  movel([0.353341, -1.417894, -2.538259, -0.756236, 1.570796, 1.924137],accel_mss,speed_ms,0,blend_radius_m)
  movel([0.350688, -1.416056, -2.539657, -0.756676, 1.570796, 1.921484],accel_mss,speed_ms,0,blend_radius_m)
  movel([0.348186, -1.414065, -2.541166, -0.757158, 1.570796, 1.918982],accel_mss,speed_ms,0,blend_radius_m)
  movel([0.345836, -1.411923, -2.542783, -0.757683, 1.570796, 1.916633],accel_mss,speed_ms,0,blend_radius_m)
  movel([0.343651, -1.409630, -2.544506, -0.758253, 1.570796, 1.914447],accel_mss,speed_ms,0,blend_radius_m)
  movel([0.342913, -1.408723, -2.545186, -0.758481, 1.570796, 1.913709],accel_mss,speed_ms,0,blend_radius_m)
  movel([0.342382, -1.407674, -2.545970, -0.758745, 1.570796, 1.913178],accel_mss,speed_ms,0,blend_radius_m)
  movel([0.342236, -1.406961, -2.546502, -0.758926, 1.570796, 1.913032],accel_mss,speed_ms,0,blend_radius_m)
  movel([0.342196, -1.406201, -2.547068, -0.759119, 1.570796, 1.912992],accel_mss,speed_ms,0,blend_radius_m)
  movel([0.342303, -1.404603, -2.548257, -0.759529, 1.570796, 1.913100],accel_mss,speed_ms,0,blend_radius_m)
  movel([0.343314, -1.398696, -2.552617, -0.761077, 1.570796, 1.914110],accel_mss,speed_ms,0,blend_radius_m)
  movel([0.343428, -1.397065, -2.553812, -0.761513, 1.570796, 1.914224],accel_mss,speed_ms,0,blend_radius_m)
  movel([0.343321, -1.395654, -2.554842, -0.761893, 1.570796, 1.914117],accel_mss,speed_ms,0,blend_radius_m)
  movel([0.343156, -1.395078, -2.555262, -0.762049, 1.570796, 1.913953],accel_mss,speed_ms,0,blend_radius_m)
  movel([0.342904, -1.394608, -2.555604, -0.762177, 1.570796, 1.913701],accel_mss,speed_ms,0,blend_radius_m)
  movel([0.342554, -1.394267, -2.555852, -0.762270, 1.570796, 1.913350],accel_mss,speed_ms,0,blend_radius_m)
  movel([0.342095, -1.394069, -2.555996, -0.762324, 1.570796, 1.912892],accel_mss,speed_ms,0,blend_radius_m)
  movel([0.341153, -1.393966, -2.556071, -0.762352, 1.570796, 1.911950],accel_mss,speed_ms,0,blend_radius_m)
  movel([0.340728, -1.393866, -2.556143, -0.762379, 1.570796, 1.911524],accel_mss,speed_ms,0,blend_radius_m)
  movel([0.340432, -1.393631, -2.556314, -0.762444, 1.570796, 1.911229],accel_mss,speed_ms,0,blend_radius_m)
  movel([0.340359, -1.393040, -2.556743, -0.762606, 1.570796, 1.911155],accel_mss,speed_ms,0,blend_radius_m)
  movel([0.340573, -1.392339, -2.557251, -0.762798, 1.570796, 1.911370],accel_mss,speed_ms,0,blend_radius_m)
  movel([0.341367, -1.390085, -2.558881, -0.763423, 1.570796, 1.912163],accel_mss,speed_ms,0,blend_radius_m)
  movel([0.342003, -1.387856, -2.560485, -0.764048, 1.570796, 1.912799],accel_mss,speed_ms,0,blend_radius_m)
  movel([0.342890, -1.383456, -2.563631, -0.765302, 1.570796, 1.913686],accel_mss,speed_ms,0,blend_radius_m)
  movel([0.343413, -1.379085, -2.566728, -0.766576, 1.570796, 1.914210],accel_mss,speed_ms,0,blend_radius_m)
  movel([0.343750, -1.374694, -2.569812, -0.767883, 1.570796, 1.914546],accel_mss,speed_ms,0,blend_radius_m)
  speed_ms = 0.005
  movel([0.343750, -1.366094, -2.565773, -0.780522, 1.570796, 1.914546],accel_mss,speed_ms,0,blend_radius_m)
  speed_ms = 0.040
  movel([0.339869, -1.373054, -2.560934, -0.778400, 1.570796, 1.910666],accel_mss,speed_ms,0,blend_radius_m)
  speed_ms = 0.005
  movel([0.339869, -1.381608, -2.564943, -0.765837, 1.570796, 1.910666],accel_mss,speed_ms,0,blend_radius_m)
  speed_ms = 0.025
  movel([0.337589, -1.386297, -2.561603, -0.764489, 1.570796, 1.908385],accel_mss,speed_ms,0,blend_radius_m)
  movel([0.336311, -1.388619, -2.559937, -0.763833, 1.570796, 1.907108],accel_mss,speed_ms,0,blend_radius_m)
  movel([0.334950, -1.390919, -2.558279, -0.763191, 1.570796, 1.905746],accel_mss,speed_ms,0,blend_radius_m)
  movel([0.333977, -1.389868, -2.559037, -0.763483, 1.570796, 1.904774],accel_mss,speed_ms,0,blend_radius_m)
  movel([0.333786, -1.389712, -2.559150, -0.763527, 1.570796, 1.904582],accel_mss,speed_ms,0,blend_radius_m)
  movel([0.333516, -1.389690, -2.559166, -0.763533, 1.570796, 1.904313],accel_mss,speed_ms,0,blend_radius_m)
  movel([0.333217, -1.389876, -2.559032, -0.763481, 1.570796, 1.904013],accel_mss,speed_ms,0,blend_radius_m)
  movel([0.332976, -1.390157, -2.558829, -0.763403, 1.570796, 1.903772],accel_mss,speed_ms,0,blend_radius_m)
  movel([0.331482, -1.391896, -2.557572, -0.762921, 1.570796, 1.902279],accel_mss,speed_ms,0,blend_radius_m)
  movel([0.329770, -1.393485, -2.556421, -0.762484, 1.570796, 1.900566],accel_mss,speed_ms,0,blend_radius_m)
  movel([0.329322, -1.393797, -2.556193, -0.762398, 1.570796, 1.900118],accel_mss,speed_ms,0,blend_radius_m)
  movel([0.328892, -1.393891, -2.556126, -0.762373, 1.570796, 1.899688],accel_mss,speed_ms,0,blend_radius_m)
  movel([0.328696, -1.393685, -2.556275, -0.762429, 1.570796, 1.899492],accel_mss,speed_ms,0,blend_radius_m)
  movel([0.328675, -1.393350, -2.556518, -0.762521, 1.570796, 1.899472],accel_mss,speed_ms,0,blend_radius_m)
  movel([0.328990, -1.391182, -2.558089, -0.763118, 1.570796, 1.899786],accel_mss,speed_ms,0,blend_radius_m)
  movel([0.329681, -1.388937, -2.559708, -0.763744, 1.570796, 1.900478],accel_mss,speed_ms,0,blend_radius_m)
  speed_ms = 0.005
  movel([0.329681, -1.380434, -2.555730, -0.776225, 1.570796, 1.900478],accel_mss,speed_ms,0,blend_radius_m)
  speed_ms = 0.040
  movel([0.332271, -1.385014, -2.552462, -0.774913, 1.570796, 1.903067],accel_mss,speed_ms,0,blend_radius_m)
  speed_ms = 0.005
  movel([0.332271, -1.393486, -2.556420, -0.762483, 1.570796, 1.903067],accel_mss,speed_ms,0,blend_radius_m)
  speed_ms = 0.025
  movel([0.331292, -1.396772, -2.554026, -0.761592, 1.570796, 1.902088],accel_mss,speed_ms,0,blend_radius_m)
  movel([0.330631, -1.398425, -2.552816, -0.761149, 1.570796, 1.901428],accel_mss,speed_ms,0,blend_radius_m)
  movel([0.328994, -1.401710, -2.550398, -0.760281, 1.570796, 1.899790],accel_mss,speed_ms,0,blend_radius_m)
  movel([0.328023, -1.403329, -2.549201, -0.759859, 1.570796, 1.898819],accel_mss,speed_ms,0,blend_radius_m)
  movel([0.325798, -1.406488, -2.546855, -0.759046, 1.570796, 1.896594],accel_mss,speed_ms,0,blend_radius_m)
  movel([0.326216, -1.405393, -2.547669, -0.759326, 1.570796, 1.897012],accel_mss,speed_ms,0,blend_radius_m)
  movel([0.326316, -1.404349, -2.548445, -0.759595, 1.570796, 1.897112],accel_mss,speed_ms,0,blend_radius_m)
  movel([0.326100, -1.403427, -2.549128, -0.759833, 1.570796, 1.896896],accel_mss,speed_ms,0,blend_radius_m)
  movel([0.325568, -1.402702, -2.549666, -0.760022, 1.570796, 1.896365],accel_mss,speed_ms,0,blend_radius_m)
  speed_ms = 0.005
  movel([0.325568, -1.394294, -2.545747, -0.772348, 1.570796, 1.896365],accel_mss,speed_ms,0,blend_radius_m)
  speed_ms = 0.040
  movel([0.312695, -1.397176, -2.543637, -0.771576, 1.570796, 1.883492],accel_mss,speed_ms,0,blend_radius_m)
  speed_ms = 0.005
  movel([0.312695, -1.405564, -2.547543, -0.759283, 1.570796, 1.883492],accel_mss,speed_ms,0,blend_radius_m)
  speed_ms = 0.025
  movel([0.310320, -1.407416, -2.546163, -0.758811, 1.570796, 1.881117],accel_mss,speed_ms,0,blend_radius_m)
  movel([0.307808, -1.409042, -2.544946, -0.758400, 1.570796, 1.878604],accel_mss,speed_ms,0,blend_radius_m)
  movel([0.305202, -1.410422, -2.543912, -0.758055, 1.570796, 1.875999],accel_mss,speed_ms,0,blend_radius_m)
  movel([0.302547, -1.411527, -2.543081, -0.757781, 1.570796, 1.873344],accel_mss,speed_ms,0,blend_radius_m)
  movel([0.303286, -1.410545, -2.543819, -0.758025, 1.570796, 1.874082],accel_mss,speed_ms,0,blend_radius_m)
  movel([0.303859, -1.409585, -2.544540, -0.758264, 1.570796, 1.874656],accel_mss,speed_ms,0,blend_radius_m)
  movel([0.304225, -1.408734, -2.545177, -0.758478, 1.570796, 1.875021],accel_mss,speed_ms,0,blend_radius_m)
  movel([0.304341, -1.408081, -2.545666, -0.758642, 1.570796, 1.875137],accel_mss,speed_ms,0,blend_radius_m)
  movel([0.304161, -1.407717, -2.545938, -0.758734, 1.570796, 1.874957],accel_mss,speed_ms,0,blend_radius_m)
  movel([0.303948, -1.407671, -2.545972, -0.758746, 1.570796, 1.874744],accel_mss,speed_ms,0,blend_radius_m)
  movel([0.303642, -1.407729, -2.545928, -0.758731, 1.570796, 1.874438],accel_mss,speed_ms,0,blend_radius_m)
  movel([0.302742, -1.408211, -2.545569, -0.758610, 1.570796, 1.873539],accel_mss,speed_ms,0,blend_radius_m)
  movel([0.300391, -1.410083, -2.544167, -0.758140, 1.570796, 1.871188],accel_mss,speed_ms,0,blend_radius_m)
  movel([0.299301, -1.410867, -2.543577, -0.757945, 1.570796, 1.870098],accel_mss,speed_ms,0,blend_radius_m)
  movel([0.296993, -1.412235, -2.542548, -0.757606, 1.570796, 1.867789],accel_mss,speed_ms,0,blend_radius_m)
  movel([0.295802, -1.412800, -2.542122, -0.757467, 1.570796, 1.866599],accel_mss,speed_ms,0,blend_radius_m)
  movel([0.294607, -1.413268, -2.541769, -0.757352, 1.570796, 1.865403],accel_mss,speed_ms,0,blend_radius_m)
  movel([0.293418, -1.413635, -2.541492, -0.757263, 1.570796, 1.864215],accel_mss,speed_ms,0,blend_radius_m)
  movel([0.292256, -1.413884, -2.541303, -0.757202, 1.570796, 1.863052],accel_mss,speed_ms,0,blend_radius_m)
  movel([0.293826, -1.412474, -2.542367, -0.757547, 1.570796, 1.864623],accel_mss,speed_ms,0,blend_radius_m)
  movel([0.295363, -1.411029, -2.543456, -0.757904, 1.570796, 1.866160],accel_mss,speed_ms,0,blend_radius_m)
  movel([0.296110, -1.409980, -2.544243, -0.758165, 1.570796, 1.866906],accel_mss,speed_ms,0,blend_radius_m)
  movel([0.296586, -1.408893, -2.545058, -0.758438, 1.570796, 1.867383],accel_mss,speed_ms,0,blend_radius_m)
  movel([0.296599, -1.408490, -2.545359, -0.758539, 1.570796, 1.867396],accel_mss,speed_ms,0,blend_radius_m)
  movel([0.296393, -1.408265, -2.545528, -0.758596, 1.570796, 1.867190],accel_mss,speed_ms,0,blend_radius_m)
  movel([0.295922, -1.408281, -2.545516, -0.758592, 1.570796, 1.866719],accel_mss,speed_ms,0,blend_radius_m)
  movel([0.295135, -1.408602, -2.545276, -0.758511, 1.570796, 1.865931],accel_mss,speed_ms,0,blend_radius_m)
  movel([0.290915, -1.410859, -2.543584, -0.757947, 1.570796, 1.861712],accel_mss,speed_ms,0,blend_radius_m)
  movel([0.288820, -1.411752, -2.542911, -0.757725, 1.570796, 1.859616],accel_mss,speed_ms,0,blend_radius_m)
  movel([0.287788, -1.412048, -2.542689, -0.757652, 1.570796, 1.858584],accel_mss,speed_ms,0,blend_radius_m)
  movel([0.286768, -1.412208, -2.542568, -0.757613, 1.570796, 1.857565],accel_mss,speed_ms,0,blend_radius_m)
  speed_ms = 0.005
  movel([0.286768, -1.403867, -2.538690, -0.769831, 1.570796, 1.857565],accel_mss,speed_ms,0,blend_radius_m)
  speed_ms = 0.040
  movel([0.307123, -1.384967, -2.552495, -0.774927, 1.570796, 1.877919],accel_mss,speed_ms,0,blend_radius_m)
  speed_ms = 0.005
  movel([0.307123, -1.393440, -2.556453, -0.762496, 1.570796, 1.877919],accel_mss,speed_ms,0,blend_radius_m)
  speed_ms = 0.025
  movel([0.307349, -1.392012, -2.557488, -0.762888, 1.570796, 1.878145],accel_mss,speed_ms,0,blend_radius_m)
  movel([0.307875, -1.390552, -2.558544, -0.763293, 1.570796, 1.878671],accel_mss,speed_ms,0,blend_radius_m)
  movel([0.308665, -1.389081, -2.559605, -0.763704, 1.570796, 1.879461],accel_mss,speed_ms,0,blend_radius_m)
  movel([0.309681, -1.387631, -2.560646, -0.764111, 1.570796, 1.880477],accel_mss,speed_ms,0,blend_radius_m)
  movel([0.310891, -1.386226, -2.561654, -0.764509, 1.570796, 1.881688],accel_mss,speed_ms,0,blend_radius_m)
  movel([0.312255, -1.384897, -2.562603, -0.764888, 1.570796, 1.883051],accel_mss,speed_ms,0,blend_radius_m)
  movel([0.313741, -1.383669, -2.563479, -0.765241, 1.570796, 1.884537],accel_mss,speed_ms,0,blend_radius_m)
  movel([0.315307, -1.382571, -2.564260, -0.765558, 1.570796, 1.886103],accel_mss,speed_ms,0,blend_radius_m)
  movel([0.317303, -1.381387, -2.565100, -0.765902, 1.570796, 1.888099],accel_mss,speed_ms,0,blend_radius_m)
  movel([0.321349, -1.379143, -2.566687, -0.766559, 1.570796, 1.892145],accel_mss,speed_ms,0,blend_radius_m)
  movel([0.323312, -1.377877, -2.567579, -0.766933, 1.570796, 1.894108],accel_mss,speed_ms,0,blend_radius_m)
  movel([0.325159, -1.376347, -2.568654, -0.767388, 1.570796, 1.895955],accel_mss,speed_ms,0,blend_radius_m)
  movel([0.325987, -1.375488, -2.569256, -0.767645, 1.570796, 1.896784],accel_mss,speed_ms,0,blend_radius_m)
  movel([0.326715, -1.374590, -2.569885, -0.767914, 1.570796, 1.897511],accel_mss,speed_ms,0,blend_radius_m)
  movel([0.327314, -1.373670, -2.570527, -0.768192, 1.570796, 1.898111],accel_mss,speed_ms,0,blend_radius_m)
  movel([0.327760, -1.372746, -2.571172, -0.768472, 1.570796, 1.898557],accel_mss,speed_ms,0,blend_radius_m)
  movel([0.328019, -1.371841, -2.571802, -0.768747, 1.570796, 1.898816],accel_mss,speed_ms,0,blend_radius_m)
  movel([0.328063, -1.370972, -2.572405, -0.769012, 1.570796, 1.898860],accel_mss,speed_ms,0,blend_radius_m)
  speed_ms = 0.005
  movel([0.328063, -1.362347, -2.568349, -0.781693, 1.570796, 1.898860],accel_mss,speed_ms,0,blend_radius_m)
  speed_ms = 0.040
  movel([0.327969, -1.355374, -2.573093, -0.783923, 1.570796, 1.898765],accel_mss,speed_ms,0,blend_radius_m)
  speed_ms = 0.005
  movel([0.327969, -1.364044, -2.577178, -0.771166, 1.570796, 1.898765],accel_mss,speed_ms,0,blend_radius_m)
  speed_ms = 0.025
  movel([0.325748, -1.369382, -2.573506, -0.769501, 1.570796, 1.896545],accel_mss,speed_ms,0,blend_radius_m)
  movel([0.325014, -1.370536, -2.572707, -0.769146, 1.570796, 1.895810],accel_mss,speed_ms,0,blend_radius_m)
  movel([0.323980, -1.371546, -2.572006, -0.768837, 1.570796, 1.894777],accel_mss,speed_ms,0,blend_radius_m)
  movel([0.322764, -1.372368, -2.571435, -0.768586, 1.570796, 1.893560],accel_mss,speed_ms,0,blend_radius_m)
  movel([0.318705, -1.374593, -2.569882, -0.767913, 1.570796, 1.889501],accel_mss,speed_ms,0,blend_radius_m)
  movel([0.317313, -1.375524, -2.569231, -0.767634, 1.570796, 1.888110],accel_mss,speed_ms,0,blend_radius_m)
  movel([0.315981, -1.376546, -2.568514, -0.767328, 1.570796, 1.886777],accel_mss,speed_ms,0,blend_radius_m)
  movel([0.314719, -1.377645, -2.567743, -0.767002, 1.570796, 1.885516],accel_mss,speed_ms,0,blend_radius_m)
  movel([0.313629, -1.378816, -2.566918, -0.766655, 1.570796, 1.884425],accel_mss,speed_ms,0,blend_radius_m)
  movel([0.312677, -1.380053, -2.566044, -0.766292, 1.570796, 1.883473],accel_mss,speed_ms,0,blend_radius_m)
  movel([0.311739, -1.381287, -2.565171, -0.765931, 1.570796, 1.882535],accel_mss,speed_ms,0,blend_radius_m)
  movel([0.310692, -1.382453, -2.564344, -0.765592, 1.570796, 1.881488],accel_mss,speed_ms,0,blend_radius_m)
  movel([0.310217, -1.379416, -2.566495, -0.766479, 1.570796, 1.881013],accel_mss,speed_ms,0,blend_radius_m)
  movel([0.310427, -1.378523, -2.567124, -0.766742, 1.570796, 1.881223],accel_mss,speed_ms,0,blend_radius_m)
  movel([0.310784, -1.377639, -2.567747, -0.767003, 1.570796, 1.881580],accel_mss,speed_ms,0,blend_radius_m)
  movel([0.311287, -1.376761, -2.568364, -0.767264, 1.570796, 1.882083],accel_mss,speed_ms,0,blend_radius_m)
  movel([0.311945, -1.375885, -2.568978, -0.767526, 1.570796, 1.882741],accel_mss,speed_ms,0,blend_radius_m)
  movel([0.313120, -1.374783, -2.569750, -0.767856, 1.570796, 1.883917],accel_mss,speed_ms,0,blend_radius_m)
  movel([0.314797, -1.373557, -2.570606, -0.768226, 1.570796, 1.885594],accel_mss,speed_ms,0,blend_radius_m)
  movel([0.318871, -1.370934, -2.572431, -0.769024, 1.570796, 1.889668],accel_mss,speed_ms,0,blend_radius_m)
  movel([0.320876, -1.369641, -2.573327, -0.769421, 1.570796, 1.891672],accel_mss,speed_ms,0,blend_radius_m)
  movel([0.322594, -1.368424, -2.574168, -0.769796, 1.570796, 1.893391],accel_mss,speed_ms,0,blend_radius_m)
  movel([0.323827, -1.367340, -2.574916, -0.770133, 1.570796, 1.894624],accel_mss,speed_ms,0,blend_radius_m)
  movel([0.324201, -1.366860, -2.575247, -0.770283, 1.570796, 1.894997],accel_mss,speed_ms,0,blend_radius_m)
  movel([0.324377, -1.366430, -2.575542, -0.770417, 1.570796, 1.895173],accel_mss,speed_ms,0,blend_radius_m)
  speed_ms = 0.005
  movel([0.324377, -1.357775, -2.571467, -0.783147, 1.570796, 1.895173],accel_mss,speed_ms,0,blend_radius_m)
  speed_ms = 0.040
  movel([0.317644, -1.355816, -2.572794, -0.783779, 1.570796, 1.888440],accel_mss,speed_ms,0,blend_radius_m)
  speed_ms = 0.005
  movel([0.317644, -1.364484, -2.576878, -0.771028, 1.570796, 1.888440],accel_mss,speed_ms,0,blend_radius_m)
  speed_ms = 0.025
  movel([0.316995, -1.364280, -2.577017, -0.771092, 1.570796, 1.887792],accel_mss,speed_ms,0,blend_radius_m)
  movel([0.316480, -1.363934, -2.577254, -0.771201, 1.570796, 1.887276],accel_mss,speed_ms,0,blend_radius_m)
  movel([0.315783, -1.362916, -2.577950, -0.771524, 1.570796, 1.886579],accel_mss,speed_ms,0,blend_radius_m)
  movel([0.315427, -1.361607, -2.578842, -0.771940, 1.570796, 1.886224],accel_mss,speed_ms,0,blend_radius_m)
  movel([0.315292, -1.360185, -2.579809, -0.772396, 1.570796, 1.886089],accel_mss,speed_ms,0,blend_radius_m)
  movel([0.315340, -1.359638, -2.580180, -0.772572, 1.570796, 1.886136],accel_mss,speed_ms,0,blend_radius_m)
  movel([0.315896, -1.358775, -2.580764, -0.772850, 1.570796, 1.886692],accel_mss,speed_ms,0,blend_radius_m)
  movel([0.317769, -1.356422, -2.582353, -0.773614, 1.570796, 1.888565],accel_mss,speed_ms,0,blend_radius_m)
  movel([0.321286, -1.351596, -2.585588, -0.775206, 1.570796, 1.892083],accel_mss,speed_ms,0,blend_radius_m)
  movel([0.322923, -1.349133, -2.587226, -0.776031, 1.570796, 1.893720],accel_mss,speed_ms,0,blend_radius_m)
  speed_ms = 0.005
  movel([0.322923, -1.340366, -2.583075, -0.788949, 1.570796, 1.893720],accel_mss,speed_ms,0,blend_radius_m)
  speed_ms = 0.040
  movel([0.318249, -1.341582, -2.582277, -0.788530, 1.570796, 1.889045],accel_mss,speed_ms,0,blend_radius_m)
  speed_ms = 0.005
  movel([0.318249, -1.350341, -2.586423, -0.775625, 1.570796, 1.889045],accel_mss,speed_ms,0,blend_radius_m)
  speed_ms = 0.025
  movel([0.317404, -1.351859, -2.585412, -0.775118, 1.570796, 1.888200],accel_mss,speed_ms,0,blend_radius_m)
  movel([0.316388, -1.353339, -2.584423, -0.774627, 1.570796, 1.887185],accel_mss,speed_ms,0,blend_radius_m)
  movel([0.315173, -1.354678, -2.583525, -0.774186, 1.570796, 1.885969],accel_mss,speed_ms,0,blend_radius_m)
  movel([0.314479, -1.355266, -2.583131, -0.773992, 1.570796, 1.885275],accel_mss,speed_ms,0,blend_radius_m)
  movel([0.312991, -1.356296, -2.582438, -0.773655, 1.570796, 1.883787],accel_mss,speed_ms,0,blend_radius_m)
  movel([0.312589, -1.356891, -2.582037, -0.773461, 1.570796, 1.883385],accel_mss,speed_ms,0,blend_radius_m)
  movel([0.310058, -1.361595, -2.578850, -0.771944, 1.570796, 1.880854],accel_mss,speed_ms,0,blend_radius_m)
  movel([0.309827, -1.362051, -2.578539, -0.771798, 1.570796, 1.880623],accel_mss,speed_ms,0,blend_radius_m)
  movel([0.309727, -1.362487, -2.578242, -0.771660, 1.570796, 1.880524],accel_mss,speed_ms,0,blend_radius_m)
  movel([0.309968, -1.362959, -2.577920, -0.771510, 1.570796, 1.880764],accel_mss,speed_ms,0,blend_radius_m)
  movel([0.310464, -1.363243, -2.577726, -0.771420, 1.570796, 1.881260],accel_mss,speed_ms,0,blend_radius_m)
  movel([0.311933, -1.363994, -2.577213, -0.771182, 1.570796, 1.882730],accel_mss,speed_ms,0,blend_radius_m)
  movel([0.313243, -1.364912, -2.576584, -0.770893, 1.570796, 1.884039],accel_mss,speed_ms,0,blend_radius_m)
  movel([0.314279, -1.366052, -2.575802, -0.770535, 1.570796, 1.885076],accel_mss,speed_ms,0,blend_radius_m)
  movel([0.314920, -1.367474, -2.574824, -0.770091, 1.570796, 1.885717],accel_mss,speed_ms,0,blend_radius_m)
  speed_ms = 0.005
  movel([0.314920, -1.358825, -2.570753, -0.782811, 1.570796, 1.885717],accel_mss,speed_ms,0,blend_radius_m)
  speed_ms = 0.040
  movel([0.308499, -1.370918, -2.562427, -0.779044, 1.570796, 1.879295],accel_mss,speed_ms,0,blend_radius_m)
  speed_ms = 0.005
  movel([0.308499, -1.379486, -2.566445, -0.766458, 1.570796, 1.879295],accel_mss,speed_ms,0,blend_radius_m)
  speed_ms = 0.025
  movel([0.308142, -1.379675, -2.566311, -0.766402, 1.570796, 1.878938],accel_mss,speed_ms,0,blend_radius_m)
  movel([0.307804, -1.379962, -2.566109, -0.766318, 1.570796, 1.878600],accel_mss,speed_ms,0,blend_radius_m)
  movel([0.306398, -1.381586, -2.564959, -0.765844, 1.570796, 1.877194],accel_mss,speed_ms,0,blend_radius_m)
  movel([0.306182, -1.381703, -2.564876, -0.765810, 1.570796, 1.876978],accel_mss,speed_ms,0,blend_radius_m)
  movel([0.305890, -1.381676, -2.564896, -0.765818, 1.570796, 1.876686],accel_mss,speed_ms,0,blend_radius_m)
  movel([0.305691, -1.381462, -2.565047, -0.765880, 1.570796, 1.876488],accel_mss,speed_ms,0,blend_radius_m)
  movel([0.305524, -1.380686, -2.565597, -0.766106, 1.570796, 1.876321],accel_mss,speed_ms,0,blend_radius_m)
  movel([0.305660, -1.379126, -2.566699, -0.766564, 1.570796, 1.876456],accel_mss,speed_ms,0,blend_radius_m)
  movel([0.306239, -1.377612, -2.567766, -0.767011, 1.570796, 1.877035],accel_mss,speed_ms,0,blend_radius_m)
  movel([0.307051, -1.376086, -2.568837, -0.767465, 1.570796, 1.877848],accel_mss,speed_ms,0,blend_radius_m)
  movel([0.307976, -1.374599, -2.569878, -0.767911, 1.570796, 1.878772],accel_mss,speed_ms,0,blend_radius_m)
  movel([0.309020, -1.373202, -2.570853, -0.768333, 1.570796, 1.879816],accel_mss,speed_ms,0,blend_radius_m)
  movel([0.310178, -1.371895, -2.571763, -0.768730, 1.570796, 1.880974],accel_mss,speed_ms,0,blend_radius_m)
  movel([0.311443, -1.370676, -2.572610, -0.769103, 1.570796, 1.882240],accel_mss,speed_ms,0,blend_radius_m)
  movel([0.312813, -1.369539, -2.573398, -0.769452, 1.570796, 1.883610],accel_mss,speed_ms,0,blend_radius_m)
  movel([0.314279, -1.368486, -2.574126, -0.769777, 1.570796, 1.885075],accel_mss,speed_ms,0,blend_radius_m)
  movel([0.315839, -1.367510, -2.574799, -0.770080, 1.570796, 1.886635],accel_mss,speed_ms,0,blend_radius_m)
  movel([0.317485, -1.366610, -2.575418, -0.770361, 1.570796, 1.888282],accel_mss,speed_ms,0,blend_radius_m)
  movel([0.319775, -1.365190, -2.576393, -0.770805, 1.570796, 1.890571],accel_mss,speed_ms,0,blend_radius_m)
  movel([0.322192, -1.363404, -2.577616, -0.771369, 1.570796, 1.892989],accel_mss,speed_ms,0,blend_radius_m)
  movel([0.324813, -1.361260, -2.579078, -0.772051, 1.570796, 1.895609],accel_mss,speed_ms,0,blend_radius_m)
  speed_ms = 0.005
  movel([0.324813, -1.352571, -2.574980, -0.784838, 1.570796, 1.895609],accel_mss,speed_ms,0,blend_radius_m)
  speed_ms = 0.040
  movel([0.322789, -1.352336, -2.575138, -0.784915, 1.570796, 1.893585],accel_mss,speed_ms,0,blend_radius_m)
  speed_ms = 0.005
  movel([0.322789, -1.361026, -2.579237, -0.772126, 1.570796, 1.893585],accel_mss,speed_ms,0,blend_radius_m)
  speed_ms = 0.025
  movel([0.325060, -1.357489, -2.581633, -0.773266, 1.570796, 1.895856],accel_mss,speed_ms,0,blend_radius_m)
  movel([0.327540, -1.353985, -2.583990, -0.774414, 1.570796, 1.898337],accel_mss,speed_ms,0,blend_radius_m)
  movel([0.328901, -1.352289, -2.585125, -0.774975, 1.570796, 1.899697],accel_mss,speed_ms,0,blend_radius_m)
  movel([0.330358, -1.350651, -2.586217, -0.775521, 1.570796, 1.901154],accel_mss,speed_ms,0,blend_radius_m)
  movel([0.331934, -1.349089, -2.587255, -0.776045, 1.570796, 1.902731],accel_mss,speed_ms,0,blend_radius_m)
  movel([0.333636, -1.347623, -2.588226, -0.776540, 1.570796, 1.904433],accel_mss,speed_ms,0,blend_radius_m)
  movel([0.338281, -1.344182, -2.590494, -0.777714, 1.570796, 1.909077],accel_mss,speed_ms,0,blend_radius_m)
  movel([0.340290, -1.342554, -2.591561, -0.778274, 1.570796, 1.911086],accel_mss,speed_ms,0,blend_radius_m)
  movel([0.341243, -1.341682, -2.592131, -0.778576, 1.570796, 1.912039],accel_mss,speed_ms,0,blend_radius_m)
  movel([0.342119, -1.340743, -2.592744, -0.778902, 1.570796, 1.912915],accel_mss,speed_ms,0,blend_radius_m)
  movel([0.344165, -1.337635, -2.594763, -0.779991, 1.570796, 1.914961],accel_mss,speed_ms,0,blend_radius_m)
  speed_ms = 0.005
  movel([0.344165, -1.328796, -2.590561, -0.793032, 1.570796, 1.914961],accel_mss,speed_ms,0,blend_radius_m)
  speed_ms = 0.040
  movel([0.349051, -1.321604, -2.595125, -0.795660, 1.570796, 1.919847],accel_mss,speed_ms,0,blend_radius_m)
  speed_ms = 0.005
  movel([0.349051, -1.330486, -2.599359, -0.782543, 1.570796, 1.919847],accel_mss,speed_ms,0,blend_radius_m)
  speed_ms = 0.025
  movel([0.350619, -1.327900, -2.601005, -0.783484, 1.570796, 1.921415],accel_mss,speed_ms,0,blend_radius_m)
  movel([0.351604, -1.326705, -2.601762, -0.783922, 1.570796, 1.922400],accel_mss,speed_ms,0,blend_radius_m)
  movel([0.352794, -1.325669, -2.602418, -0.784303, 1.570796, 1.923590],accel_mss,speed_ms,0,blend_radius_m)
  movel([0.353735, -1.325094, -2.602780, -0.784515, 1.570796, 1.924531],accel_mss,speed_ms,0,blend_radius_m)
  movel([0.354708, -1.324645, -2.603064, -0.784681, 1.570796, 1.925504],accel_mss,speed_ms,0,blend_radius_m)
  movel([0.356688, -1.323931, -2.603513, -0.784945, 1.570796, 1.927484],accel_mss,speed_ms,0,blend_radius_m)
  movel([0.358468, -1.323146, -2.604007, -0.785236, 1.570796, 1.929265],accel_mss,speed_ms,0,blend_radius_m)
  movel([0.359922, -1.322182, -2.604612, -0.785595, 1.570796, 1.930719],accel_mss,speed_ms,0,blend_radius_m)
  movel([0.362751, -1.319636, -2.606203, -0.786549, 1.570796, 1.933547],accel_mss,speed_ms,0,blend_radius_m)
  movel([0.363357, -1.319157, -2.606502, -0.786730, 1.570796, 1.934153],accel_mss,speed_ms,0,blend_radius_m)
  movel([0.364004, -1.318782, -2.606736, -0.786871, 1.570796, 1.934800],accel_mss,speed_ms,0,blend_radius_m)
  movel([0.365382, -1.318258, -2.607061, -0.787069, 1.570796, 1.936179],accel_mss,speed_ms,0,blend_radius_m)
  movel([0.368164, -1.317488, -2.607540, -0.787361, 1.570796, 1.938960],accel_mss,speed_ms,0,blend_radius_m)
  movel([0.371123, -1.316378, -2.608228, -0.787783, 1.570796, 1.941919],accel_mss,speed_ms,0,blend_radius_m)
  movel([0.372596, -1.315685, -2.608657, -0.788047, 1.570796, 1.943392],accel_mss,speed_ms,0,blend_radius_m)
  movel([0.374034, -1.314815, -2.609194, -0.788379, 1.570796, 1.944830],accel_mss,speed_ms,0,blend_radius_m)
  movel([0.375107, -1.313914, -2.609750, -0.788725, 1.570796, 1.945903],accel_mss,speed_ms,0,blend_radius_m)
  movel([0.375975, -1.312857, -2.610400, -0.789131, 1.570796, 1.946771],accel_mss,speed_ms,0,blend_radius_m)
  movel([0.376436, -1.311818, -2.611038, -0.789533, 1.570796, 1.947232],accel_mss,speed_ms,0,blend_radius_m)
  movel([0.376451, -1.311361, -2.611318, -0.789709, 1.570796, 1.947248],accel_mss,speed_ms,0,blend_radius_m)
  movel([0.376289, -1.310975, -2.611555, -0.789859, 1.570796, 1.947085],accel_mss,speed_ms,0,blend_radius_m)
  movel([0.375621, -1.310415, -2.611897, -0.790077, 1.570796, 1.946417],accel_mss,speed_ms,0,blend_radius_m)
  movel([0.374663, -1.310045, -2.612124, -0.790220, 1.570796, 1.945460],accel_mss,speed_ms,0,blend_radius_m)
  movel([0.373483, -1.309859, -2.612237, -0.790293, 1.570796, 1.944279],accel_mss,speed_ms,0,blend_radius_m)
  movel([0.372161, -1.309843, -2.612247, -0.790299, 1.570796, 1.942958],accel_mss,speed_ms,0,blend_radius_m)
  movel([0.370770, -1.309993, -2.612155, -0.790241, 1.570796, 1.941566],accel_mss,speed_ms,0,blend_radius_m)
  movel([0.369387, -1.310295, -2.611971, -0.790123, 1.570796, 1.940183],accel_mss,speed_ms,0,blend_radius_m)
  movel([0.368086, -1.310742, -2.611697, -0.789950, 1.570796, 1.938882],accel_mss,speed_ms,0,blend_radius_m)
  movel([0.366941, -1.311323, -2.611342, -0.789724, 1.570796, 1.937738],accel_mss,speed_ms,0,blend_radius_m)
  movel([0.365361, -1.312504, -2.610617, -0.789268, 1.570796, 1.936157],accel_mss,speed_ms,0,blend_radius_m)
  movel([0.360899, -1.316398, -2.608216, -0.787775, 1.570796, 1.931696],accel_mss,speed_ms,0,blend_radius_m)
  movel([0.357794, -1.318784, -2.606735, -0.786871, 1.570796, 1.928590],accel_mss,speed_ms,0,blend_radius_m)
  movel([0.354959, -1.320535, -2.605642, -0.786211, 1.570796, 1.925755],accel_mss,speed_ms,0,blend_radius_m)
  movel([0.353550, -1.321372, -2.605119, -0.785898, 1.570796, 1.924347],accel_mss,speed_ms,0,blend_radius_m)
  movel([0.352205, -1.322311, -2.604531, -0.785547, 1.570796, 1.923002],accel_mss,speed_ms,0,blend_radius_m)
  movel([0.350915, -1.323430, -2.603828, -0.785131, 1.570796, 1.921711],accel_mss,speed_ms,0,blend_radius_m)
  movel([0.349740, -1.324629, -2.603073, -0.784686, 1.570796, 1.920536],accel_mss,speed_ms,0,blend_radius_m)
  movel([0.348669, -1.325894, -2.602275, -0.784220, 1.570796, 1.919466],accel_mss,speed_ms,0,blend_radius_m)
  movel([0.347691, -1.327204, -2.601446, -0.783739, 1.570796, 1.918487],accel_mss,speed_ms,0,blend_radius_m)
  movel([0.345956, -1.329897, -2.599735, -0.782757, 1.570796, 1.916752],accel_mss,speed_ms,0,blend_radius_m)
  movel([0.344424, -1.332576, -2.598023, -0.781790, 1.570796, 1.915221],accel_mss,speed_ms,0,blend_radius_m)
  speed_ms = 0.005
  movel([0.344424, -1.323706, -2.593798, -0.794885, 1.570796, 1.915221],accel_mss,speed_ms,0,blend_radius_m)
  speed_ms = 0.040
  movel([0.340785, -1.325157, -2.592879, -0.794353, 1.570796, 1.911581],accel_mss,speed_ms,0,blend_radius_m)
  speed_ms = 0.005
  movel([0.340785, -1.334019, -2.597097, -0.781273, 1.570796, 1.911581],accel_mss,speed_ms,0,blend_radius_m)
  speed_ms = 0.025
  movel([0.343327, -1.329820, -2.599784, -0.782785, 1.570796, 1.914124],accel_mss,speed_ms,0,blend_radius_m)
  movel([0.344465, -1.328079, -2.600891, -0.783419, 1.570796, 1.915261],accel_mss,speed_ms,0,blend_radius_m)
  movel([0.345507, -1.326318, -2.602007, -0.784064, 1.570796, 1.916304],accel_mss,speed_ms,0,blend_radius_m)
  movel([0.346218, -1.324778, -2.602980, -0.784631, 1.570796, 1.917014],accel_mss,speed_ms,0,blend_radius_m)
  movel([0.346717, -1.323245, -2.603944, -0.785199, 1.570796, 1.917514],accel_mss,speed_ms,0,blend_radius_m)
  movel([0.346996, -1.321750, -2.604882, -0.785757, 1.570796, 1.917792],accel_mss,speed_ms,0,blend_radius_m)
  movel([0.347046, -1.320325, -2.605774, -0.786290, 1.570796, 1.917842],accel_mss,speed_ms,0,blend_radius_m)
  movel([0.347778, -1.320120, -2.605901, -0.786367, 1.570796, 1.918574],accel_mss,speed_ms,0,blend_radius_m)
  movel([0.348472, -1.320081, -2.605926, -0.786382, 1.570796, 1.919268],accel_mss,speed_ms,0,blend_radius_m)
  movel([0.349799, -1.320203, -2.605850, -0.786336, 1.570796, 1.920596],accel_mss,speed_ms,0,blend_radius_m)
  movel([0.351211, -1.320202, -2.605850, -0.786337, 1.570796, 1.922008],accel_mss,speed_ms,0,blend_radius_m)
  movel([0.351944, -1.320017, -2.605966, -0.786406, 1.570796, 1.922741],accel_mss,speed_ms,0,blend_radius_m)
  movel([0.352658, -1.319621, -2.606213, -0.786555, 1.570796, 1.923455],accel_mss,speed_ms,0,blend_radius_m)
  movel([0.360769, -1.313713, -2.609874, -0.788802, 1.570796, 1.931565],accel_mss,speed_ms,0,blend_radius_m)
  movel([0.360914, -1.312683, -2.610507, -0.789199, 1.570796, 1.931710],accel_mss,speed_ms,0,blend_radius_m)
  movel([0.360736, -1.311745, -2.611083, -0.789561, 1.570796, 1.931532],accel_mss,speed_ms,0,blend_radius_m)
  movel([0.360245, -1.310950, -2.611570, -0.789869, 1.570796, 1.931041],accel_mss,speed_ms,0,blend_radius_m)
  movel([0.359461, -1.310345, -2.611940, -0.790104, 1.570796, 1.930257],accel_mss,speed_ms,0,blend_radius_m)
  movel([0.361095, -1.310189, -2.612035, -0.790164, 1.570796, 1.931891],accel_mss,speed_ms,0,blend_radius_m)
  movel([0.362585, -1.310328, -2.611951, -0.790110, 1.570796, 1.933381],accel_mss,speed_ms,0,blend_radius_m)
  movel([0.363857, -1.310746, -2.611695, -0.789948, 1.570796, 1.934653],accel_mss,speed_ms,0,blend_radius_m)
  movel([0.364841, -1.311428, -2.611277, -0.789684, 1.570796, 1.935638],accel_mss,speed_ms,0,blend_radius_m)
  speed_ms = 0.005
  movel([0.364841, -1.302433, -2.606958, -0.802997, 1.570796, 1.935638],accel_mss,speed_ms,0,blend_radius_m)
  speed_ms = 0.040
  movel([0.366450, -1.298436, -2.609366, -0.804587, 1.570796, 1.937246],accel_mss,speed_ms,0,blend_radius_m)
  speed_ms = 0.005
  movel([0.366450, -1.307453, -2.613703, -0.791233, 1.570796, 1.937246],accel_mss,speed_ms,0,blend_radius_m)
  speed_ms = 0.025
  movel([0.367612, -1.305388, -2.614955, -0.792046, 1.570796, 1.938409],accel_mss,speed_ms,0,blend_radius_m)
  movel([0.368567, -1.303391, -2.616160, -0.792838, 1.570796, 1.939363],accel_mss,speed_ms,0,blend_radius_m)
  movel([0.369330, -1.301451, -2.617326, -0.793612, 1.570796, 1.940127],accel_mss,speed_ms,0,blend_radius_m)
  movel([0.369916, -1.299553, -2.618462, -0.794374, 1.570796, 1.940712],accel_mss,speed_ms,0,blend_radius_m)
  movel([0.370339, -1.297683, -2.619577, -0.795129, 1.570796, 1.941136],accel_mss,speed_ms,0,blend_radius_m)
  movel([0.370616, -1.295823, -2.620681, -0.795885, 1.570796, 1.941412],accel_mss,speed_ms,0,blend_radius_m)
  movel([0.370788, -1.292081, -2.622890, -0.797419, 1.570796, 1.941585],accel_mss,speed_ms,0,blend_radius_m)
  movel([0.366939, -1.299226, -2.618657, -0.794506, 1.570796, 1.937735],accel_mss,speed_ms,0,blend_radius_m)
  movel([0.367292, -1.298430, -2.619132, -0.794827, 1.570796, 1.938088],accel_mss,speed_ms,0,blend_radius_m)
  movel([0.367497, -1.297648, -2.619598, -0.795144, 1.570796, 1.938293],accel_mss,speed_ms,0,blend_radius_m)
  movel([0.367519, -1.296136, -2.620495, -0.795757, 1.570796, 1.938316],accel_mss,speed_ms,0,blend_radius_m)
  movel([0.367103, -1.294716, -2.621336, -0.796337, 1.570796, 1.937900],accel_mss,speed_ms,0,blend_radius_m)
  movel([0.366356, -1.293414, -2.622105, -0.796870, 1.570796, 1.937153],accel_mss,speed_ms,0,blend_radius_m)
  movel([0.365380, -1.292252, -2.622789, -0.797348, 1.570796, 1.936177],accel_mss,speed_ms,0,blend_radius_m)
  movel([0.364283, -1.291257, -2.623373, -0.797759, 1.570796, 1.935079],accel_mss,speed_ms,0,blend_radius_m)
  movel([0.362143, -1.289862, -2.624190, -0.798336, 1.570796, 1.932940],accel_mss,speed_ms,0,blend_radius_m)
  movel([0.362715, -1.292997, -2.622350, -0.797042, 1.570796, 1.933512],accel_mss,speed_ms,0,blend_radius_m)
  movel([0.362706, -1.294725, -2.621331, -0.796333, 1.570796, 1.933502],accel_mss,speed_ms,0,blend_radius_m)
  movel([0.362303, -1.296437, -2.620317, -0.795635, 1.570796, 1.933099],accel_mss,speed_ms,0,blend_radius_m)
  movel([0.361334, -1.296243, -2.620432, -0.795714, 1.570796, 1.932130],accel_mss,speed_ms,0,blend_radius_m)
  movel([0.360464, -1.295867, -2.620655, -0.795867, 1.570796, 1.931260],accel_mss,speed_ms,0,blend_radius_m)
  movel([0.358870, -1.294799, -2.621287, -0.796303, 1.570796, 1.929667],accel_mss,speed_ms,0,blend_radius_m)
  movel([0.357242, -1.293700, -2.621936, -0.796753, 1.570796, 1.928038],accel_mss,speed_ms,0,blend_radius_m)
  movel([0.356327, -1.293283, -2.622182, -0.796924, 1.570796, 1.927123],accel_mss,speed_ms,0,blend_radius_m)
  movel([0.355301, -1.293031, -2.622330, -0.797027, 1.570796, 1.926098],accel_mss,speed_ms,0,blend_radius_m)
  movel([0.354062, -1.294848, -2.621258, -0.796283, 1.570796, 1.924858],accel_mss,speed_ms,0,blend_radius_m)
  movel([0.353191, -1.296710, -2.620155, -0.795524, 1.570796, 1.923987],accel_mss,speed_ms,0,blend_radius_m)
  movel([0.351729, -1.296578, -2.620233, -0.795578, 1.570796, 1.922525],accel_mss,speed_ms,0,blend_radius_m)
  movel([0.350418, -1.296205, -2.620455, -0.795729, 1.570796, 1.921214],accel_mss,speed_ms,0,blend_radius_m)
  movel([0.349284, -1.295596, -2.620816, -0.795978, 1.570796, 1.920081],accel_mss,speed_ms,0,blend_radius_m)
  movel([0.348362, -1.294767, -2.621306, -0.796316, 1.570796, 1.919158],accel_mss,speed_ms,0,blend_radius_m)
  movel([0.348169, -1.294931, -2.621209, -0.796249, 1.570796, 1.918966],accel_mss,speed_ms,0,blend_radius_m)
  movel([0.346493, -1.297166, -2.619884, -0.795339, 1.570796, 1.917289],accel_mss,speed_ms,0,blend_radius_m)
  movel([0.344537, -1.299992, -2.618199, -0.794197, 1.570796, 1.915334],accel_mss,speed_ms,0,blend_radius_m)
  movel([0.343774, -1.301395, -2.617359, -0.793634, 1.570796, 1.914570],accel_mss,speed_ms,0,blend_radius_m)
  movel([0.343191, -1.302708, -2.616571, -0.793110, 1.570796, 1.913987],accel_mss,speed_ms,0,blend_radius_m)
  movel([0.342295, -1.305435, -2.614926, -0.792028, 1.570796, 1.913091],accel_mss,speed_ms,0,blend_radius_m)
  movel([0.339280, -1.301953, -2.617025, -0.793411, 1.570796, 1.910076],accel_mss,speed_ms,0,blend_radius_m)
  movel([0.338412, -1.303418, -2.616144, -0.792827, 1.570796, 1.909208],accel_mss,speed_ms,0,blend_radius_m)
  movel([0.337665, -1.304909, -2.615244, -0.792236, 1.570796, 1.908461],accel_mss,speed_ms,0,blend_radius_m)
  movel([0.336498, -1.307921, -2.613419, -0.791050, 1.570796, 1.907295],accel_mss,speed_ms,0,blend_radius_m)
  movel([0.335736, -1.310876, -2.611615, -0.789898, 1.570796, 1.906533],accel_mss,speed_ms,0,blend_radius_m)
  movel([0.335196, -1.314520, -2.609376, -0.788492, 1.570796, 1.905992],accel_mss,speed_ms,0,blend_radius_m)
  movel([0.335024, -1.314949, -2.609112, -0.788328, 1.570796, 1.905820],accel_mss,speed_ms,0,blend_radius_m)
  movel([0.334735, -1.315355, -2.608861, -0.788173, 1.570796, 1.905531],accel_mss,speed_ms,0,blend_radius_m)
  movel([0.334180, -1.315791, -2.608591, -0.788006, 1.570796, 1.904976],accel_mss,speed_ms,0,blend_radius_m)
  movel([0.330116, -1.317718, -2.607397, -0.787274, 1.570796, 1.900913],accel_mss,speed_ms,0,blend_radius_m)
  movel([0.328059, -1.318419, -2.606962, -0.787009, 1.570796, 1.898855],accel_mss,speed_ms,0,blend_radius_m)
  movel([0.327318, -1.318499, -2.606912, -0.786978, 1.570796, 1.898114],accel_mss,speed_ms,0,blend_radius_m)
  movel([0.326909, -1.318306, -2.607032, -0.787051, 1.570796, 1.897705],accel_mss,speed_ms,0,blend_radius_m)
  movel([0.328384, -1.320291, -2.605795, -0.786303, 1.570796, 1.899180],accel_mss,speed_ms,0,blend_radius_m)
  movel([0.329282, -1.321145, -2.605261, -0.785983, 1.570796, 1.900078],accel_mss,speed_ms,0,blend_radius_m)
  movel([0.330278, -1.321902, -2.604787, -0.785700, 1.570796, 1.901074],accel_mss,speed_ms,0,blend_radius_m)
  movel([0.326692, -1.324729, -2.603010, -0.784649, 1.570796, 1.897488],accel_mss,speed_ms,0,blend_radius_m)
  movel([0.322877, -1.327949, -2.600974, -0.783466, 1.570796, 1.893673],accel_mss,speed_ms,0,blend_radius_m)
  movel([0.321056, -1.329646, -2.599895, -0.782848, 1.570796, 1.891852],accel_mss,speed_ms,0,blend_radius_m)
  movel([0.319382, -1.331364, -2.598798, -0.782226, 1.570796, 1.890178],accel_mss,speed_ms,0,blend_radius_m)
  movel([0.317925, -1.333083, -2.597698, -0.781608, 1.570796, 1.888721],accel_mss,speed_ms,0,blend_radius_m)
  movel([0.316752, -1.334773, -2.596611, -0.781004, 1.570796, 1.887548],accel_mss,speed_ms,0,blend_radius_m)
  movel([0.318428, -1.333869, -2.597193, -0.781327, 1.570796, 1.889225],accel_mss,speed_ms,0,blend_radius_m)
  movel([0.320123, -1.333125, -2.597671, -0.781593, 1.570796, 1.890919],accel_mss,speed_ms,0,blend_radius_m)
  movel([0.321814, -1.332566, -2.598029, -0.781794, 1.570796, 1.892610],accel_mss,speed_ms,0,blend_radius_m)
  movel([0.323490, -1.332214, -2.598255, -0.781920, 1.570796, 1.894287],accel_mss,speed_ms,0,blend_radius_m)
  movel([0.322315, -1.333028, -2.597733, -0.781628, 1.570796, 1.893111],accel_mss,speed_ms,0,blend_radius_m)
  movel([0.320130, -1.334873, -2.596547, -0.780969, 1.570796, 1.890927],accel_mss,speed_ms,0,blend_radius_m)
  movel([0.319137, -1.335888, -2.595893, -0.780608, 1.570796, 1.889933],accel_mss,speed_ms,0,blend_radius_m)
  movel([0.317396, -1.338040, -2.594501, -0.779848, 1.570796, 1.888192],accel_mss,speed_ms,0,blend_radius_m)
  movel([0.316664, -1.339162, -2.593773, -0.779454, 1.570796, 1.887460],accel_mss,speed_ms,0,blend_radius_m)
  movel([0.316038, -1.340298, -2.593034, -0.779057, 1.570796, 1.886834],accel_mss,speed_ms,0,blend_radius_m)
  speed_ms = 0.005
  movel([0.316038, -1.331475, -2.588843, -0.792070, 1.570796, 1.886834],accel_mss,speed_ms,0,blend_radius_m)
  speed_ms = 0.040
  movel([0.321417, -1.335052, -2.586535, -0.790802, 1.570796, 1.892213],accel_mss,speed_ms,0,blend_radius_m)
  speed_ms = 0.005
  movel([0.321417, -1.343852, -2.590710, -0.777827, 1.570796, 1.892213],accel_mss,speed_ms,0,blend_radius_m)
  speed_ms = 0.025
  movel([0.321926, -1.342288, -2.591735, -0.778366, 1.570796, 1.892722],accel_mss,speed_ms,0,blend_radius_m)
  movel([0.322579, -1.340695, -2.592775, -0.778919, 1.570796, 1.893375],accel_mss,speed_ms,0,blend_radius_m)
  movel([0.323372, -1.339091, -2.593819, -0.779479, 1.570796, 1.894168],accel_mss,speed_ms,0,blend_radius_m)
  movel([0.324297, -1.337496, -2.594853, -0.780040, 1.570796, 1.895094],accel_mss,speed_ms,0,blend_radius_m)
  movel([0.325354, -1.335923, -2.595870, -0.780596, 1.570796, 1.896151],accel_mss,speed_ms,0,blend_radius_m)
  movel([0.326535, -1.334390, -2.596858, -0.781141, 1.570796, 1.897331],accel_mss,speed_ms,0,blend_radius_m)
  movel([0.327833, -1.332912, -2.597807, -0.781670, 1.570796, 1.898630],accel_mss,speed_ms,0,blend_radius_m)
  movel([0.329246, -1.331509, -2.598706, -0.782174, 1.570796, 1.900042],accel_mss,speed_ms,0,blend_radius_m)
  movel([0.333839, -1.327296, -2.601388, -0.783705, 1.570796, 1.904635],accel_mss,speed_ms,0,blend_radius_m)
  movel([0.334794, -1.326250, -2.602050, -0.784089, 1.570796, 1.905590],accel_mss,speed_ms,0,blend_radius_m)
  movel([0.335665, -1.325123, -2.602762, -0.784504, 1.570796, 1.906461],accel_mss,speed_ms,0,blend_radius_m)
  movel([0.336448, -1.323877, -2.603547, -0.784965, 1.570796, 1.907244],accel_mss,speed_ms,0,blend_radius_m)
  movel([0.337143, -1.322465, -2.604434, -0.785490, 1.570796, 1.907939],accel_mss,speed_ms,0,blend_radius_m)
  movel([0.338700, -1.318362, -2.606997, -0.787030, 1.570796, 1.909497],accel_mss,speed_ms,0,blend_radius_m)
  movel([0.339578, -1.316314, -2.608268, -0.787807, 1.570796, 1.910374],accel_mss,speed_ms,0,blend_radius_m)
  movel([0.340747, -1.314285, -2.609522, -0.788583, 1.570796, 1.911544],accel_mss,speed_ms,0,blend_radius_m)
  movel([0.341642, -1.313099, -2.610252, -0.789038, 1.570796, 1.912439],accel_mss,speed_ms,0,blend_radius_m)
  movel([0.342650, -1.311973, -2.610944, -0.789473, 1.570796, 1.913446],accel_mss,speed_ms,0,blend_radius_m)
  movel([0.344931, -1.309885, -2.612221, -0.790283, 1.570796, 1.915728],accel_mss,speed_ms,0,blend_radius_m)
  movel([0.347440, -1.307973, -2.613387, -0.791030, 1.570796, 1.918236],accel_mss,speed_ms,0,blend_radius_m)
  movel([0.350033, -1.306187, -2.614471, -0.791731, 1.570796, 1.920829],accel_mss,speed_ms,0,blend_radius_m)
  movel([0.352569, -1.304534, -2.615471, -0.792384, 1.570796, 1.923365],accel_mss,speed_ms,0,blend_radius_m)
  movel([0.355169, -1.303068, -2.616355, -0.792967, 1.570796, 1.925965],accel_mss,speed_ms,0,blend_radius_m)
  movel([0.356460, -1.302481, -2.616707, -0.793200, 1.570796, 1.927257],accel_mss,speed_ms,0,blend_radius_m)
  movel([0.357735, -1.302031, -2.616978, -0.793380, 1.570796, 1.928531],accel_mss,speed_ms,0,blend_radius_m)
  movel([0.358971, -1.301752, -2.617145, -0.793492, 1.570796, 1.929767],accel_mss,speed_ms,0,blend_radius_m)
  movel([0.360166, -1.301669, -2.617195, -0.793525, 1.570796, 1.930962],accel_mss,speed_ms,0,blend_radius_m)
  speed_ms = 0.005
  movel([0.360166, -1.292619, -2.612833, -0.806937, 1.570796, 1.930962],accel_mss,speed_ms,0,blend_radius_m)
  speed_ms = 0.040
  movel([0.361313, -1.294015, -2.612004, -0.806369, 1.570796, 1.932109],accel_mss,speed_ms,0,blend_radius_m)
  speed_ms = 0.005
  movel([0.361313, -1.303057, -2.616361, -0.792971, 1.570796, 1.932109],accel_mss,speed_ms,0,blend_radius_m)
  speed_ms = 0.025
  movel([0.361689, -1.303435, -2.616134, -0.792821, 1.570796, 1.932485],accel_mss,speed_ms,0,blend_radius_m)
  movel([0.362166, -1.304074, -2.615748, -0.792567, 1.570796, 1.932962],accel_mss,speed_ms,0,blend_radius_m)
  movel([0.362734, -1.305865, -2.614666, -0.791858, 1.570796, 1.933530],accel_mss,speed_ms,0,blend_radius_m)
  movel([0.362826, -1.306873, -2.614055, -0.791461, 1.570796, 1.933622],accel_mss,speed_ms,0,blend_radius_m)
  movel([0.362721, -1.307389, -2.613741, -0.791258, 1.570796, 1.933517],accel_mss,speed_ms,0,blend_radius_m)
  movel([0.362582, -1.307494, -2.613678, -0.791217, 1.570796, 1.933379],accel_mss,speed_ms,0,blend_radius_m)
  movel([0.362364, -1.307438, -2.613712, -0.791239, 1.570796, 1.933160],accel_mss,speed_ms,0,blend_radius_m)
  movel([0.360333, -1.306108, -2.614519, -0.791762, 1.570796, 1.931129],accel_mss,speed_ms,0,blend_radius_m)
  movel([0.359138, -1.305653, -2.614794, -0.791942, 1.570796, 1.929934],accel_mss,speed_ms,0,blend_radius_m)
  movel([0.358453, -1.305583, -2.614836, -0.791969, 1.570796, 1.929250],accel_mss,speed_ms,0,blend_radius_m)
  movel([0.357695, -1.305651, -2.614795, -0.791943, 1.570796, 1.928491],accel_mss,speed_ms,0,blend_radius_m)
  movel([0.356795, -1.305916, -2.614635, -0.791838, 1.570796, 1.927592],accel_mss,speed_ms,0,blend_radius_m)
  movel([0.355885, -1.306311, -2.614396, -0.791682, 1.570796, 1.926682],accel_mss,speed_ms,0,blend_radius_m)
  movel([0.353659, -1.307485, -2.613683, -0.791221, 1.570796, 1.924455],accel_mss,speed_ms,0,blend_radius_m)
  movel([0.351448, -1.308869, -2.612841, -0.790679, 1.570796, 1.922244],accel_mss,speed_ms,0,blend_radius_m)
  movel([0.349319, -1.310419, -2.611895, -0.790075, 1.570796, 1.920115],accel_mss,speed_ms,0,blend_radius_m)
  movel([0.347345, -1.312082, -2.610876, -0.789431, 1.570796, 1.918142],accel_mss,speed_ms,0,blend_radius_m)
  movel([0.348059, -1.314542, -2.609363, -0.788484, 1.570796, 1.918856],accel_mss,speed_ms,0,blend_radius_m)
  movel([0.348419, -1.317182, -2.607730, -0.787477, 1.570796, 1.919215],accel_mss,speed_ms,0,blend_radius_m)
  movel([0.347668, -1.316638, -2.608067, -0.787684, 1.570796, 1.918464],accel_mss,speed_ms,0,blend_radius_m)
  movel([0.346749, -1.316288, -2.608284, -0.787817, 1.570796, 1.917545],accel_mss,speed_ms,0,blend_radius_m)
  movel([0.345689, -1.316149, -2.608370, -0.787870, 1.570796, 1.916485],accel_mss,speed_ms,0,blend_radius_m)
  movel([0.344526, -1.316223, -2.608324, -0.787842, 1.570796, 1.915322],accel_mss,speed_ms,0,blend_radius_m)
  movel([0.343945, -1.316449, -2.608184, -0.787756, 1.570796, 1.914742],accel_mss,speed_ms,0,blend_radius_m)
  movel([0.343645, -1.316913, -2.607897, -0.787579, 1.570796, 1.914441],accel_mss,speed_ms,0,blend_radius_m)
  movel([0.341484, -1.322083, -2.604674, -0.785632, 1.570796, 1.912280],accel_mss,speed_ms,0,blend_radius_m)
  movel([0.340185, -1.324693, -2.603033, -0.784663, 1.570796, 1.910981],accel_mss,speed_ms,0,blend_radius_m)
  movel([0.338680, -1.327322, -2.601372, -0.783696, 1.570796, 1.909477],accel_mss,speed_ms,0,blend_radius_m)
  movel([0.336985, -1.329894, -2.599737, -0.782758, 1.570796, 1.907782],accel_mss,speed_ms,0,blend_radius_m)
  movel([0.335106, -1.332340, -2.598174, -0.781875, 1.570796, 1.905903],accel_mss,speed_ms,0,blend_radius_m)
  movel([0.331165, -1.337182, -2.595056, -0.780150, 1.570796, 1.901962],accel_mss,speed_ms,0,blend_radius_m)
  movel([0.329470, -1.339649, -2.593456, -0.779284, 1.570796, 1.900266],accel_mss,speed_ms,0,blend_radius_m)
  movel([0.328120, -1.342213, -2.591784, -0.778392, 1.570796, 1.898916],accel_mss,speed_ms,0,blend_radius_m)
  speed_ms = 0.005
  movel([0.328120, -1.333402, -2.587602, -0.791385, 1.570796, 1.898916],accel_mss,speed_ms,0,blend_radius_m)
  speed_ms = 0.040
  movel([0.340510, -1.330473, -2.589487, -0.792429, 1.570796, 1.911306],accel_mss,speed_ms,0,blend_radius_m)
  speed_ms = 0.005
  movel([0.340510, -1.339302, -2.593682, -0.779405, 1.570796, 1.911306],accel_mss,speed_ms,0,blend_radius_m)
  speed_ms = 0.025
  movel([0.339440, -1.341372, -2.592333, -0.778684, 1.570796, 1.910236],accel_mss,speed_ms,0,blend_radius_m)
  movel([0.338038, -1.343382, -2.591019, -0.777989, 1.570796, 1.908834],accel_mss,speed_ms,0,blend_radius_m)
  movel([0.336354, -1.345264, -2.589782, -0.777343, 1.570796, 1.907151],accel_mss,speed_ms,0,blend_radius_m)
  movel([0.334442, -1.346961, -2.588663, -0.776764, 1.570796, 1.905238],accel_mss,speed_ms,0,blend_radius_m)
  speed_ms = 0.005
  movel([0.334442, -1.338181, -2.584502, -0.789706, 1.570796, 1.905238],accel_mss,speed_ms,0,blend_radius_m)
  speed_ms = 0.040
  movel([0.332455, -1.335199, -2.586440, -0.790750, 1.570796, 1.903251],accel_mss,speed_ms,0,blend_radius_m)
  speed_ms = 0.005
  movel([0.332455, -1.343998, -2.590614, -0.777777, 1.570796, 1.903251],accel_mss,speed_ms,0,blend_radius_m)
  speed_ms = 0.025
  movel([0.322417, -1.356103, -2.582568, -0.773718, 1.570796, 1.893214],accel_mss,speed_ms,0,blend_radius_m)
  movel([0.321897, -1.356910, -2.582024, -0.773455, 1.570796, 1.892693],accel_mss,speed_ms,0,blend_radius_m)
  movel([0.321852, -1.357860, -2.581383, -0.773146, 1.570796, 1.892648],accel_mss,speed_ms,0,blend_radius_m)
  movel([0.321791, -1.359086, -2.580554, -0.772749, 1.570796, 1.892587],accel_mss,speed_ms,0,blend_radius_m)
  movel([0.321417, -1.360387, -2.579672, -0.772331, 1.570796, 1.892213],accel_mss,speed_ms,0,blend_radius_m)
  speed_ms = 0.005
  movel([0.321417, -1.351692, -2.575570, -0.785127, 1.570796, 1.892213],accel_mss,speed_ms,0,blend_radius_m)
  speed_ms = 0.040
  movel([0.335946, -1.346058, -2.579324, -0.787006, 1.570796, 1.906742],accel_mss,speed_ms,0,blend_radius_m)
  speed_ms = 0.005
  movel([0.335946, -1.354789, -2.583451, -0.774149, 1.570796, 1.906742],accel_mss,speed_ms,0,blend_radius_m)
  speed_ms = 0.025
  movel([0.336376, -1.353408, -2.584377, -0.774604, 1.570796, 1.907173],accel_mss,speed_ms,0,blend_radius_m)
  movel([0.336990, -1.352010, -2.585311, -0.775068, 1.570796, 1.907787],accel_mss,speed_ms,0,blend_radius_m)
  movel([0.337775, -1.350620, -2.586237, -0.775531, 1.570796, 1.908572],accel_mss,speed_ms,0,blend_radius_m)
  movel([0.338725, -1.349258, -2.587143, -0.775988, 1.570796, 1.909521],accel_mss,speed_ms,0,blend_radius_m)
  movel([0.339478, -1.348347, -2.587747, -0.776295, 1.570796, 1.910275],accel_mss,speed_ms,0,blend_radius_m)
  movel([0.340322, -1.347486, -2.588317, -0.776587, 1.570796, 1.911118],accel_mss,speed_ms,0,blend_radius_m)
  movel([0.341247, -1.346723, -2.588821, -0.776846, 1.570796, 1.912043],accel_mss,speed_ms,0,blend_radius_m)
  movel([0.342256, -1.346099, -2.589232, -0.777058, 1.570796, 1.913052],accel_mss,speed_ms,0,blend_radius_m)
  movel([0.343132, -1.345754, -2.589459, -0.777175, 1.570796, 1.913928],accel_mss,speed_ms,0,blend_radius_m)
  movel([0.344055, -1.345576, -2.589577, -0.777236, 1.570796, 1.914851],accel_mss,speed_ms,0,blend_radius_m)
  movel([0.344999, -1.345533, -2.589605, -0.777251, 1.570796, 1.915795],accel_mss,speed_ms,0,blend_radius_m)
  movel([0.345946, -1.345598, -2.589562, -0.777229, 1.570796, 1.916743],accel_mss,speed_ms,0,blend_radius_m)
  movel([0.347756, -1.345924, -2.589347, -0.777117, 1.570796, 1.918552],accel_mss,speed_ms,0,blend_radius_m)
  movel([0.349306, -1.346323, -2.589085, -0.776982, 1.570796, 1.920102],accel_mss,speed_ms,0,blend_radius_m)
  movel([0.348200, -1.346151, -2.589198, -0.777040, 1.570796, 1.918996],accel_mss,speed_ms,0,blend_radius_m)
  movel([0.347008, -1.346202, -2.589164, -0.777023, 1.570796, 1.917804],accel_mss,speed_ms,0,blend_radius_m)
  movel([0.345749, -1.346506, -2.588964, -0.776919, 1.570796, 1.916545],accel_mss,speed_ms,0,blend_radius_m)
  movel([0.344437, -1.347095, -2.588575, -0.776719, 1.570796, 1.915234],accel_mss,speed_ms,0,blend_radius_m)
  movel([0.343346, -1.347820, -2.588095, -0.776473, 1.570796, 1.914142],accel_mss,speed_ms,0,blend_radius_m)
  movel([0.342338, -1.348677, -2.587528, -0.776184, 1.570796, 1.913134],accel_mss,speed_ms,0,blend_radius_m)
  movel([0.341455, -1.349566, -2.586938, -0.775885, 1.570796, 1.912251],accel_mss,speed_ms,0,blend_radius_m)
  movel([0.340669, -1.350509, -2.586311, -0.775569, 1.570796, 1.911465],accel_mss,speed_ms,0,blend_radius_m)
  movel([0.339380, -1.352505, -2.584980, -0.774903, 1.570796, 1.910176],accel_mss,speed_ms,0,blend_radius_m)
  movel([0.338455, -1.354560, -2.583604, -0.774224, 1.570796, 1.909251],accel_mss,speed_ms,0,blend_radius_m)
  movel([0.337842, -1.356748, -2.582134, -0.773508, 1.570796, 1.908638],accel_mss,speed_ms,0,blend_radius_m)
  speed_ms = 0.005
  movel([0.337842, -1.348029, -2.578016, -0.786344, 1.570796, 1.908638],accel_mss,speed_ms,0,blend_radius_m)
  speed_ms = 0.040
  movel([0.342085, -1.343604, -2.580946, -0.787838, 1.570796, 1.912881],accel_mss,speed_ms,0,blend_radius_m)
  speed_ms = 0.005
  movel([0.342085, -1.352351, -2.585083, -0.774955, 1.570796, 1.912881],accel_mss,speed_ms,0,blend_radius_m)
  speed_ms = 0.025
  movel([0.341846, -1.352648, -2.584885, -0.774856, 1.570796, 1.912643],accel_mss,speed_ms,0,blend_radius_m)
  movel([0.341486, -1.352740, -2.584823, -0.774825, 1.570796, 1.912282],accel_mss,speed_ms,0,blend_radius_m)
  movel([0.341308, -1.352548, -2.584952, -0.774889, 1.570796, 1.912105],accel_mss,speed_ms,0,blend_radius_m)
  movel([0.341343, -1.352219, -2.585171, -0.774998, 1.570796, 1.912140],accel_mss,speed_ms,0,blend_radius_m)
  movel([0.341844, -1.351571, -2.585604, -0.775214, 1.570796, 1.912640],accel_mss,speed_ms,0,blend_radius_m)
  movel([0.342154, -1.351344, -2.585755, -0.775290, 1.570796, 1.912950],accel_mss,speed_ms,0,blend_radius_m)
  movel([0.342462, -1.351357, -2.585747, -0.775285, 1.570796, 1.913258],accel_mss,speed_ms,0,blend_radius_m)
  movel([0.342582, -1.351602, -2.585583, -0.775204, 1.570796, 1.913379],accel_mss,speed_ms,0,blend_radius_m)
  movel([0.342307, -1.352269, -2.585138, -0.774982, 1.570796, 1.913103],accel_mss,speed_ms,0,blend_radius_m)
  speed_ms = 0.005
  movel([0.342307, -1.343522, -2.581000, -0.787866, 1.570796, 1.913103],accel_mss,speed_ms,0,blend_radius_m)
  speed_ms = 0.040
  movel([0.340244, -1.352325, -2.575145, -0.784919, 1.570796, 1.911040],accel_mss,speed_ms,0,blend_radius_m)
  speed_ms = 0.005
  movel([0.340244, -1.361016, -2.579244, -0.772129, 1.570796, 1.911040],accel_mss,speed_ms,0,blend_radius_m)
  speed_ms = 0.025
  movel([0.341561, -1.359981, -2.579947, -0.772461, 1.570796, 1.912358],accel_mss,speed_ms,0,blend_radius_m)
  movel([0.342706, -1.358850, -2.580714, -0.772826, 1.570796, 1.913502],accel_mss,speed_ms,0,blend_radius_m)
  movel([0.345000, -1.356566, -2.582256, -0.773567, 1.570796, 1.915797],accel_mss,speed_ms,0,blend_radius_m)
  movel([0.346861, -1.355146, -2.583211, -0.774032, 1.570796, 1.917657],accel_mss,speed_ms,0,blend_radius_m)
  movel([0.352929, -1.351242, -2.585823, -0.775324, 1.570796, 1.923725],accel_mss,speed_ms,0,blend_radius_m)
  movel([0.354104, -1.350307, -2.586446, -0.775636, 1.570796, 1.924900],accel_mss,speed_ms,0,blend_radius_m)
  movel([0.354518, -1.349777, -2.586798, -0.775814, 1.570796, 1.925314],accel_mss,speed_ms,0,blend_radius_m)
  movel([0.354676, -1.349240, -2.587154, -0.775994, 1.570796, 1.925472],accel_mss,speed_ms,0,blend_radius_m)
  movel([0.354441, -1.348728, -2.587494, -0.776167, 1.570796, 1.925237],accel_mss,speed_ms,0,blend_radius_m)
  movel([0.353935, -1.348411, -2.587704, -0.776274, 1.570796, 1.924731],accel_mss,speed_ms,0,blend_radius_m)
  movel([0.353074, -1.348088, -2.587918, -0.776383, 1.570796, 1.923870],accel_mss,speed_ms,0,blend_radius_m)
  movel([0.352170, -1.347992, -2.587981, -0.776415, 1.570796, 1.922967],accel_mss,speed_ms,0,blend_radius_m)
  movel([0.351157, -1.348137, -2.587886, -0.776366, 1.570796, 1.921953],accel_mss,speed_ms,0,blend_radius_m)
  movel([0.349972, -1.348533, -2.587623, -0.776233, 1.570796, 1.920768],accel_mss,speed_ms,0,blend_radius_m)
  movel([0.348688, -1.349169, -2.587202, -0.776018, 1.570796, 1.919484],accel_mss,speed_ms,0,blend_radius_m)
  movel([0.347408, -1.350003, -2.586648, -0.775738, 1.570796, 1.918204],accel_mss,speed_ms,0,blend_radius_m)
  movel([0.346148, -1.350985, -2.585995, -0.775410, 1.570796, 1.916944],accel_mss,speed_ms,0,blend_radius_m)
  movel([0.344920, -1.352076, -2.585267, -0.775046, 1.570796, 1.915716],accel_mss,speed_ms,0,blend_radius_m)
  movel([0.342631, -1.354390, -2.583719, -0.774280, 1.570796, 1.913427],accel_mss,speed_ms,0,blend_radius_m)
  movel([0.340658, -1.356581, -2.582246, -0.773562, 1.570796, 1.911454],accel_mss,speed_ms,0,blend_radius_m)
  movel([0.337142, -1.360701, -2.579458, -0.772230, 1.570796, 1.907938],accel_mss,speed_ms,0,blend_radius_m)
  movel([0.335890, -1.362013, -2.578565, -0.771811, 1.570796, 1.906686],accel_mss,speed_ms,0,blend_radius_m)
  movel([0.334521, -1.363249, -2.577722, -0.771418, 1.570796, 1.905317],accel_mss,speed_ms,0,blend_radius_m)
  movel([0.333037, -1.364342, -2.576974, -0.771072, 1.570796, 1.903834],accel_mss,speed_ms,0,blend_radius_m)
  movel([0.331482, -1.365212, -2.576379, -0.770799, 1.570796, 1.902279],accel_mss,speed_ms,0,blend_radius_m)
  movel([0.329898, -1.365777, -2.575991, -0.770621, 1.570796, 1.900694],accel_mss,speed_ms,0,blend_radius_m)
  movel([0.331024, -1.365802, -2.575974, -0.770613, 1.570796, 1.901820],accel_mss,speed_ms,0,blend_radius_m)
  movel([0.332200, -1.365705, -2.576040, -0.770644, 1.570796, 1.902996],accel_mss,speed_ms,0,blend_radius_m)
  movel([0.333416, -1.365485, -2.576191, -0.770713, 1.570796, 1.904212],accel_mss,speed_ms,0,blend_radius_m)
  movel([0.334651, -1.365148, -2.576423, -0.770819, 1.570796, 1.905448],accel_mss,speed_ms,0,blend_radius_m)
  movel([0.334307, -1.366444, -2.575532, -0.770412, 1.570796, 1.905103],accel_mss,speed_ms,0,blend_radius_m)
  movel([0.333751, -1.367759, -2.574627, -0.770003, 1.570796, 1.904547],accel_mss,speed_ms,0,blend_radius_m)
  movel([0.333000, -1.369061, -2.573729, -0.769600, 1.570796, 1.903797],accel_mss,speed_ms,0,blend_radius_m)
  movel([0.332072, -1.370318, -2.572859, -0.769213, 1.570796, 1.902868],accel_mss,speed_ms,0,blend_radius_m)
  movel([0.333568, -1.369228, -2.573613, -0.769548, 1.570796, 1.904364],accel_mss,speed_ms,0,blend_radius_m)
  movel([0.334934, -1.368015, -2.574450, -0.769923, 1.570796, 1.905731],accel_mss,speed_ms,0,blend_radius_m)
  movel([0.336178, -1.366699, -2.575357, -0.770333, 1.570796, 1.906974],accel_mss,speed_ms,0,blend_radius_m)
  movel([0.337312, -1.365299, -2.576319, -0.770771, 1.570796, 1.908108],accel_mss,speed_ms,0,blend_radius_m)
  movel([0.337130, -1.366165, -2.575724, -0.770500, 1.570796, 1.907926],accel_mss,speed_ms,0,blend_radius_m)
  movel([0.336729, -1.367132, -2.575059, -0.770198, 1.570796, 1.907525],accel_mss,speed_ms,0,blend_radius_m)
  movel([0.334229, -1.371430, -2.572087, -0.768872, 1.570796, 1.905025],accel_mss,speed_ms,0,blend_radius_m)
  movel([0.333706, -1.372481, -2.571356, -0.768552, 1.570796, 1.904502],accel_mss,speed_ms,0,blend_radius_m)
  movel([0.333354, -1.373467, -2.570669, -0.768253, 1.570796, 1.904151],accel_mss,speed_ms,0,blend_radius_m)
  movel([0.334394, -1.372019, -2.571678, -0.768693, 1.570796, 1.905191],accel_mss,speed_ms,0,blend_radius_m)
  movel([0.335495, -1.370711, -2.572586, -0.769092, 1.570796, 1.906291],accel_mss,speed_ms,0,blend_radius_m)
  movel([0.337832, -1.368369, -2.574206, -0.769814, 1.570796, 1.908628],accel_mss,speed_ms,0,blend_radius_m)
  movel([0.340283, -1.366127, -2.575750, -0.770512, 1.570796, 1.911079],accel_mss,speed_ms,0,blend_radius_m)
  movel([0.342774, -1.363665, -2.577438, -0.771286, 1.570796, 1.913570],accel_mss,speed_ms,0,blend_radius_m)
  movel([0.344137, -1.362034, -2.578551, -0.771804, 1.570796, 1.914933],accel_mss,speed_ms,0,blend_radius_m)
  movel([0.344998, -1.361172, -2.579138, -0.772079, 1.570796, 1.915794],accel_mss,speed_ms,0,blend_radius_m)
  movel([0.345396, -1.360889, -2.579330, -0.772170, 1.570796, 1.916192],accel_mss,speed_ms,0,blend_radius_m)
  movel([0.345747, -1.360764, -2.579415, -0.772210, 1.570796, 1.916543],accel_mss,speed_ms,0,blend_radius_m)
  movel([0.346025, -1.360817, -2.579379, -0.772193, 1.570796, 1.916821],accel_mss,speed_ms,0,blend_radius_m)
  movel([0.346226, -1.361014, -2.579246, -0.772130, 1.570796, 1.917022],accel_mss,speed_ms,0,blend_radius_m)
  movel([0.346421, -1.361690, -2.578785, -0.771914, 1.570796, 1.917218],accel_mss,speed_ms,0,blend_radius_m)
  movel([0.346364, -1.362503, -2.578231, -0.771655, 1.570796, 1.917160],accel_mss,speed_ms,0,blend_radius_m)
  movel([0.346084, -1.363166, -2.577779, -0.771444, 1.570796, 1.916881],accel_mss,speed_ms,0,blend_radius_m)
  movel([0.347604, -1.361019, -2.579242, -0.772128, 1.570796, 1.918400],accel_mss,speed_ms,0,blend_radius_m)
  movel([0.348897, -1.358811, -2.580740, -0.772838, 1.570796, 1.919693],accel_mss,speed_ms,0,blend_radius_m)
  movel([0.349949, -1.356575, -2.582250, -0.773564, 1.570796, 1.920745],accel_mss,speed_ms,0,blend_radius_m)
  movel([0.350741, -1.354340, -2.583752, -0.774297, 1.570796, 1.921538],accel_mss,speed_ms,0,blend_radius_m)
  speed_ms = 0.005
  movel([0.350741, -1.345606, -2.579624, -0.787159, 1.570796, 1.921538],accel_mss,speed_ms,0,blend_radius_m)
  speed_ms = 0.040
  movel([0.352768, -1.346714, -2.578890, -0.786785, 1.570796, 1.923565],accel_mss,speed_ms,0,blend_radius_m)
  speed_ms = 0.005
  movel([0.352768, -1.355441, -2.583013, -0.773935, 1.570796, 1.923565],accel_mss,speed_ms,0,blend_radius_m)
  speed_ms = 0.025
  movel([0.353997, -1.355953, -2.582669, -0.773767, 1.570796, 1.924793],accel_mss,speed_ms,0,blend_radius_m)
  movel([0.354409, -1.356380, -2.582381, -0.773628, 1.570796, 1.925205],accel_mss,speed_ms,0,blend_radius_m)
  movel([0.354559, -1.356975, -2.581980, -0.773434, 1.570796, 1.925355],accel_mss,speed_ms,0,blend_radius_m)
  movel([0.354437, -1.357588, -2.581567, -0.773234, 1.570796, 1.925233],accel_mss,speed_ms,0,blend_radius_m)
  movel([0.350083, -1.367866, -2.574554, -0.769970, 1.570796, 1.920879],accel_mss,speed_ms,0,blend_radius_m)
  movel([0.349730, -1.368593, -2.574052, -0.769744, 1.570796, 1.920526],accel_mss,speed_ms,0,blend_radius_m)
  movel([0.349265, -1.369302, -2.573562, -0.769525, 1.570796, 1.920062],accel_mss,speed_ms,0,blend_radius_m)
  movel([0.348684, -1.369878, -2.573163, -0.769348, 1.570796, 1.919480],accel_mss,speed_ms,0,blend_radius_m)
  movel([0.347989, -1.370208, -2.572935, -0.769247, 1.570796, 1.918785],accel_mss,speed_ms,0,blend_radius_m)
  movel([0.347380, -1.370205, -2.572937, -0.769247, 1.570796, 1.918176],accel_mss,speed_ms,0,blend_radius_m)
  movel([0.346313, -1.369849, -2.573183, -0.769357, 1.570796, 1.917109],accel_mss,speed_ms,0,blend_radius_m)
  movel([0.345700, -1.369875, -2.573165, -0.769349, 1.570796, 1.916496],accel_mss,speed_ms,0,blend_radius_m)
  movel([0.344915, -1.370293, -2.572876, -0.769220, 1.570796, 1.915711],accel_mss,speed_ms,0,blend_radius_m)
  movel([0.344180, -1.370889, -2.572462, -0.769038, 1.570796, 1.914976],accel_mss,speed_ms,0,blend_radius_m)
  movel([0.343269, -1.371526, -2.572020, -0.768843, 1.570796, 1.914065],accel_mss,speed_ms,0,blend_radius_m)
  movel([0.342306, -1.372017, -2.571678, -0.768693, 1.570796, 1.913102],accel_mss,speed_ms,0,blend_radius_m)
  movel([0.341327, -1.372358, -2.571442, -0.768589, 1.570796, 1.912124],accel_mss,speed_ms,0,blend_radius_m)
  movel([0.340365, -1.372544, -2.571312, -0.768533, 1.570796, 1.911161],accel_mss,speed_ms,0,blend_radius_m)
  movel([0.339450, -1.372574, -2.571291, -0.768524, 1.570796, 1.910247],accel_mss,speed_ms,0,blend_radius_m)
  movel([0.338624, -1.372440, -2.571385, -0.768565, 1.570796, 1.909420],accel_mss,speed_ms,0,blend_radius_m)
  movel([0.337914, -1.372144, -2.571590, -0.768655, 1.570796, 1.908710],accel_mss,speed_ms,0,blend_radius_m)
  movel([0.337358, -1.371675, -2.571917, -0.768798, 1.570796, 1.908154],accel_mss,speed_ms,0,blend_radius_m)
  speed_ms = 0.005
  movel([0.337358, -1.363054, -2.567865, -0.781470, 1.570796, 1.908154],accel_mss,speed_ms,0,blend_radius_m)
  speed_ms = 0.040
  movel([0.328691, -1.371761, -2.561839, -0.778789, 1.570796, 1.899488],accel_mss,speed_ms,0,blend_radius_m)
  speed_ms = 0.005
  movel([0.328691, -1.380323, -2.565853, -0.766212, 1.570796, 1.899488],accel_mss,speed_ms,0,blend_radius_m)
  speed_ms = 0.025
  movel([0.326379, -1.390249, -2.558763, -0.763377, 1.570796, 1.897176],accel_mss,speed_ms,0,blend_radius_m)
  movel([0.325969, -1.391472, -2.557879, -0.763038, 1.570796, 1.896765],accel_mss,speed_ms,0,blend_radius_m)
  movel([0.325601, -1.392042, -2.557467, -0.762880, 1.570796, 1.896397],accel_mss,speed_ms,0,blend_radius_m)
  movel([0.325075, -1.392518, -2.557122, -0.762749, 1.570796, 1.895871],accel_mss,speed_ms,0,blend_radius_m)
  movel([0.323725, -1.393260, -2.556584, -0.762545, 1.570796, 1.894521],accel_mss,speed_ms,0,blend_radius_m)
  movel([0.323254, -1.393847, -2.556157, -0.762385, 1.570796, 1.894050],accel_mss,speed_ms,0,blend_radius_m)
  movel([0.323014, -1.394496, -2.555685, -0.762208, 1.570796, 1.893810],accel_mss,speed_ms,0,blend_radius_m)
  movel([0.322947, -1.395526, -2.554935, -0.761928, 1.570796, 1.893743],accel_mss,speed_ms,0,blend_radius_m)
  movel([0.323169, -1.396485, -2.554235, -0.761669, 1.570796, 1.893966],accel_mss,speed_ms,0,blend_radius_m)
  movel([0.323833, -1.398248, -2.552945, -0.761196, 1.570796, 1.894630],accel_mss,speed_ms,0,blend_radius_m)
  movel([0.324019, -1.399532, -2.552003, -0.760854, 1.570796, 1.894816],accel_mss,speed_ms,0,blend_radius_m)
  movel([0.323999, -1.401451, -2.550590, -0.760349, 1.570796, 1.894795],accel_mss,speed_ms,0,blend_radius_m)
  movel([0.323818, -1.402347, -2.549927, -0.760114, 1.570796, 1.894614],accel_mss,speed_ms,0,blend_radius_m)
  movel([0.323470, -1.403049, -2.549409, -0.759931, 1.570796, 1.894267],accel_mss,speed_ms,0,blend_radius_m)
  movel([0.323222, -1.403286, -2.549233, -0.759870, 1.570796, 1.894019],accel_mss,speed_ms,0,blend_radius_m)
  movel([0.322919, -1.403431, -2.549126, -0.759832, 1.570796, 1.893716],accel_mss,speed_ms,0,blend_radius_m)
  movel([0.322556, -1.403469, -2.549098, -0.759823, 1.570796, 1.893352],accel_mss,speed_ms,0,blend_radius_m)
  movel([0.322129, -1.403381, -2.549162, -0.759845, 1.570796, 1.892925],accel_mss,speed_ms,0,blend_radius_m)
  movel([0.321841, -1.404145, -2.548596, -0.759647, 1.570796, 1.892637],accel_mss,speed_ms,0,blend_radius_m)
  movel([0.321736, -1.404996, -2.547964, -0.759428, 1.570796, 1.892532],accel_mss,speed_ms,0,blend_radius_m)
  movel([0.321919, -1.406817, -2.546609, -0.758963, 1.570796, 1.892716],accel_mss,speed_ms,0,blend_radius_m)
  movel([0.322389, -1.408543, -2.545320, -0.758526, 1.570796, 1.893185],accel_mss,speed_ms,0,blend_radius_m)
  movel([0.322861, -1.409877, -2.544321, -0.758191, 1.570796, 1.893657],accel_mss,speed_ms,0,blend_radius_m)
  movel([0.323615, -1.411230, -2.543304, -0.757854, 1.570796, 1.894411],accel_mss,speed_ms,0,blend_radius_m)
  movel([0.324564, -1.412538, -2.542319, -0.757531, 1.570796, 1.895361],accel_mss,speed_ms,0,blend_radius_m)
  movel([0.325295, -1.413946, -2.541256, -0.757187, 1.570796, 1.896091],accel_mss,speed_ms,0,blend_radius_m)
  movel([0.325450, -1.414729, -2.540663, -0.756996, 1.570796, 1.896246],accel_mss,speed_ms,0,blend_radius_m)
  movel([0.325394, -1.415590, -2.540011, -0.756788, 1.570796, 1.896191],accel_mss,speed_ms,0,blend_radius_m)
  movel([0.325234, -1.416059, -2.539655, -0.756675, 1.570796, 1.896030],accel_mss,speed_ms,0,blend_radius_m)
  movel([0.324943, -1.416518, -2.539306, -0.756564, 1.570796, 1.895739],accel_mss,speed_ms,0,blend_radius_m)
  movel([0.324560, -1.416865, -2.539043, -0.756481, 1.570796, 1.895357],accel_mss,speed_ms,0,blend_radius_m)
  movel([0.324119, -1.416998, -2.538941, -0.756449, 1.570796, 1.894915],accel_mss,speed_ms,0,blend_radius_m)
  movel([0.323820, -1.416904, -2.539013, -0.756472, 1.570796, 1.894617],accel_mss,speed_ms,0,blend_radius_m)
  movel([0.323607, -1.416707, -2.539163, -0.756519, 1.570796, 1.894403],accel_mss,speed_ms,0,blend_radius_m)
  movel([0.321948, -1.414520, -2.540822, -0.757047, 1.570796, 1.892744],accel_mss,speed_ms,0,blend_radius_m)
  movel([0.321264, -1.413319, -2.541730, -0.757340, 1.570796, 1.892060],accel_mss,speed_ms,0,blend_radius_m)
  movel([0.320685, -1.412048, -2.542688, -0.757652, 1.570796, 1.891481],accel_mss,speed_ms,0,blend_radius_m)
  movel([0.320275, -1.412468, -2.542372, -0.757549, 1.570796, 1.891071],accel_mss,speed_ms,0,blend_radius_m)
  movel([0.319969, -1.412932, -2.542022, -0.757435, 1.570796, 1.890765],accel_mss,speed_ms,0,blend_radius_m)
  movel([0.319635, -1.413962, -2.541244, -0.757183, 1.570796, 1.890432],accel_mss,speed_ms,0,blend_radius_m)
  movel([0.319604, -1.415080, -2.540398, -0.756911, 1.570796, 1.890400],accel_mss,speed_ms,0,blend_radius_m)
  movel([0.319804, -1.416225, -2.539529, -0.756635, 1.570796, 1.890600],accel_mss,speed_ms,0,blend_radius_m)
  movel([0.320575, -1.418382, -2.537887, -0.756120, 1.570796, 1.891372],accel_mss,speed_ms,0,blend_radius_m)
  movel([0.321343, -1.419972, -2.536673, -0.755744, 1.570796, 1.892139],accel_mss,speed_ms,0,blend_radius_m)
  movel([0.321549, -1.420603, -2.536189, -0.755596, 1.570796, 1.892346],accel_mss,speed_ms,0,blend_radius_m)
  movel([0.321523, -1.420951, -2.535923, -0.755515, 1.570796, 1.892319],accel_mss,speed_ms,0,blend_radius_m)
  movel([0.321340, -1.421311, -2.535647, -0.755431, 1.570796, 1.892137],accel_mss,speed_ms,0,blend_radius_m)
  movel([0.321003, -1.421647, -2.535389, -0.755353, 1.570796, 1.891800],accel_mss,speed_ms,0,blend_radius_m)
  movel([0.320672, -1.421806, -2.535267, -0.755316, 1.570796, 1.891468],accel_mss,speed_ms,0,blend_radius_m)
  movel([0.320041, -1.421782, -2.535285, -0.755321, 1.570796, 1.890838],accel_mss,speed_ms,0,blend_radius_m)
  movel([0.319197, -1.421648, -2.535388, -0.755353, 1.570796, 1.889993],accel_mss,speed_ms,0,blend_radius_m)
  movel([0.318953, -1.421777, -2.535290, -0.755323, 1.570796, 1.889749],accel_mss,speed_ms,0,blend_radius_m)
  movel([0.318707, -1.422089, -2.535049, -0.755250, 1.570796, 1.889503],accel_mss,speed_ms,0,blend_radius_m)
  movel([0.318572, -1.422466, -2.534760, -0.755163, 1.570796, 1.889368],accel_mss,speed_ms,0,blend_radius_m)
  movel([0.318555, -1.423322, -2.534101, -0.754966, 1.570796, 1.889351],accel_mss,speed_ms,0,blend_radius_m)
  movel([0.318879, -1.424801, -2.532961, -0.754627, 1.570796, 1.889675],accel_mss,speed_ms,0,blend_radius_m)
  movel([0.319795, -1.427821, -2.530621, -0.753946, 1.570796, 1.890592],accel_mss,speed_ms,0,blend_radius_m)
  movel([0.320783, -1.430790, -2.528308, -0.753290, 1.570796, 1.891580],accel_mss,speed_ms,0,blend_radius_m)
  movel([0.320879, -1.431436, -2.527803, -0.753149, 1.570796, 1.891675],accel_mss,speed_ms,0,blend_radius_m)
  movel([0.320814, -1.432137, -2.527255, -0.752997, 1.570796, 1.891610],accel_mss,speed_ms,0,blend_radius_m)
  movel([0.320517, -1.432796, -2.526739, -0.752855, 1.570796, 1.891313],accel_mss,speed_ms,0,blend_radius_m)
  movel([0.320264, -1.433079, -2.526517, -0.752794, 1.570796, 1.891061],accel_mss,speed_ms,0,blend_radius_m)
  movel([0.319579, -1.433460, -2.526217, -0.752712, 1.570796, 1.890375],accel_mss,speed_ms,0,blend_radius_m)
  movel([0.319254, -1.433512, -2.526177, -0.752701, 1.570796, 1.890050],accel_mss,speed_ms,0,blend_radius_m)
  movel([0.318675, -1.433382, -2.526279, -0.752728, 1.570796, 1.889472],accel_mss,speed_ms,0,blend_radius_m)
  movel([0.318202, -1.433040, -2.526547, -0.752802, 1.570796, 1.888998],accel_mss,speed_ms,0,blend_radius_m)
  movel([0.317845, -1.432593, -2.526898, -0.752898, 1.570796, 1.888641],accel_mss,speed_ms,0,blend_radius_m)
  movel([0.316122, -1.429688, -2.529168, -0.753532, 1.570796, 1.886918],accel_mss,speed_ms,0,blend_radius_m)
  movel([0.314590, -1.426643, -2.531535, -0.754210, 1.570796, 1.885386],accel_mss,speed_ms,0,blend_radius_m)
  movel([0.313260, -1.423461, -2.533994, -0.754934, 1.570796, 1.884057],accel_mss,speed_ms,0,blend_radius_m)
  movel([0.312137, -1.420146, -2.536539, -0.755703, 1.570796, 1.882933],accel_mss,speed_ms,0,blend_radius_m)
  movel([0.311808, -1.418870, -2.537515, -0.756004, 1.570796, 1.882604],accel_mss,speed_ms,0,blend_radius_m)
  movel([0.311719, -1.417494, -2.538564, -0.756331, 1.570796, 1.882515],accel_mss,speed_ms,0,blend_radius_m)
  movel([0.311853, -1.416621, -2.539228, -0.756540, 1.570796, 1.882649],accel_mss,speed_ms,0,blend_radius_m)
  movel([0.312103, -1.415727, -2.539907, -0.756755, 1.570796, 1.882899],accel_mss,speed_ms,0,blend_radius_m)
  movel([0.312796, -1.413906, -2.541287, -0.757197, 1.570796, 1.883593],accel_mss,speed_ms,0,blend_radius_m)
  movel([0.315929, -1.407344, -2.546216, -0.758829, 1.570796, 1.886725],accel_mss,speed_ms,0,blend_radius_m)
  movel([0.316650, -1.405481, -2.547604, -0.759304, 1.570796, 1.887446],accel_mss,speed_ms,0,blend_radius_m)
  movel([0.317084, -1.403805, -2.548848, -0.759735, 1.570796, 1.887881],accel_mss,speed_ms,0,blend_radius_m)
  movel([0.317157, -1.403081, -2.549385, -0.759923, 1.570796, 1.887953],accel_mss,speed_ms,0,blend_radius_m)
  movel([0.317106, -1.402457, -2.549846, -0.760085, 1.570796, 1.887902],accel_mss,speed_ms,0,blend_radius_m)
  movel([0.316920, -1.401950, -2.550221, -0.760218, 1.570796, 1.887717],accel_mss,speed_ms,0,blend_radius_m)
  movel([0.316584, -1.401578, -2.550496, -0.760315, 1.570796, 1.887380],accel_mss,speed_ms,0,blend_radius_m)
  movel([0.315774, -1.401161, -2.550804, -0.760425, 1.570796, 1.886570],accel_mss,speed_ms,0,blend_radius_m)
  movel([0.315429, -1.400912, -2.550987, -0.760490, 1.570796, 1.886226],accel_mss,speed_ms,0,blend_radius_m)
  movel([0.315252, -1.400546, -2.551256, -0.760586, 1.570796, 1.886048],accel_mss,speed_ms,0,blend_radius_m)
  movel([0.315411, -1.399831, -2.551783, -0.760775, 1.570796, 1.886207],accel_mss,speed_ms,0,blend_radius_m)
  movel([0.315872, -1.399080, -2.552335, -0.760974, 1.570796, 1.886668],accel_mss,speed_ms,0,blend_radius_m)
  movel([0.317443, -1.396693, -2.554084, -0.761613, 1.570796, 1.888240],accel_mss,speed_ms,0,blend_radius_m)
  movel([0.318867, -1.394288, -2.555837, -0.762264, 1.570796, 1.889663],accel_mss,speed_ms,0,blend_radius_m)
  movel([0.320164, -1.391861, -2.557598, -0.762930, 1.570796, 1.890960],accel_mss,speed_ms,0,blend_radius_m)
  movel([0.321354, -1.389413, -2.559366, -0.763611, 1.570796, 1.892150],accel_mss,speed_ms,0,blend_radius_m)
  movel([0.323510, -1.384455, -2.562919, -0.765015, 1.570796, 1.894306],accel_mss,speed_ms,0,blend_radius_m)
  movel([0.325511, -1.379405, -2.566502, -0.766482, 1.570796, 1.896307],accel_mss,speed_ms,0,blend_radius_m)
  speed_ms = 0.005
  movel([0.325511, -1.370836, -2.562484, -0.779069, 1.570796, 1.896307],accel_mss,speed_ms,0,blend_radius_m)
  speed_ms = 0.040
  movel([0.318291, -1.383265, -2.553713, -0.775410, 1.570796, 1.889087],accel_mss,speed_ms,0,blend_radius_m)
  speed_ms = 0.005
  movel([0.318291, -1.391750, -2.557678, -0.762961, 1.570796, 1.889087],accel_mss,speed_ms,0,blend_radius_m)
  speed_ms = 0.025
  movel([0.314967, -1.394440, -2.555726, -0.762223, 1.570796, 1.885764],accel_mss,speed_ms,0,blend_radius_m)
  movel([0.311570, -1.397005, -2.553855, -0.761529, 1.570796, 1.882366],accel_mss,speed_ms,0,blend_radius_m)
  movel([0.308105, -1.399445, -2.552066, -0.760878, 1.570796, 1.878901],accel_mss,speed_ms,0,blend_radius_m)
  movel([0.304585, -1.401750, -2.550369, -0.760270, 1.570796, 1.875381],accel_mss,speed_ms,0,blend_radius_m)
  movel([0.307412, -1.399037, -2.552366, -0.760986, 1.570796, 1.878208],accel_mss,speed_ms,0,blend_radius_m)
  movel([0.310073, -1.396188, -2.554452, -0.761749, 1.570796, 1.880870],accel_mss,speed_ms,0,blend_radius_m)
  movel([0.312550, -1.393221, -2.556612, -0.762556, 1.570796, 1.883347],accel_mss,speed_ms,0,blend_radius_m)
  movel([0.314826, -1.390155, -2.558830, -0.763403, 1.570796, 1.885623],accel_mss,speed_ms,0,blend_radius_m)
  movel([0.312032, -1.392337, -2.557253, -0.762799, 1.570796, 1.882828],accel_mss,speed_ms,0,blend_radius_m)
  movel([0.309185, -1.394423, -2.555739, -0.762228, 1.570796, 1.879981],accel_mss,speed_ms,0,blend_radius_m)
  movel([0.306285, -1.396410, -2.554290, -0.761689, 1.570796, 1.877082],accel_mss,speed_ms,0,blend_radius_m)
  movel([0.303342, -1.398292, -2.552912, -0.761184, 1.570796, 1.874138],accel_mss,speed_ms,0,blend_radius_m)
  movel([0.300044, -1.400314, -2.551427, -0.760648, 1.570796, 1.870840],accel_mss,speed_ms,0,blend_radius_m)
  movel([0.296845, -1.402481, -2.549829, -0.760079, 1.570796, 1.867641],accel_mss,speed_ms,0,blend_radius_m)
  movel([0.295336, -1.403703, -2.548924, -0.759762, 1.570796, 1.866132],accel_mss,speed_ms,0,blend_radius_m)
  movel([0.293946, -1.405032, -2.547938, -0.759419, 1.570796, 1.864742],accel_mss,speed_ms,0,blend_radius_m)
  movel([0.292745, -1.406454, -2.546880, -0.759055, 1.570796, 1.863541],accel_mss,speed_ms,0,blend_radius_m)
  movel([0.291792, -1.407948, -2.545765, -0.758676, 1.570796, 1.862588],accel_mss,speed_ms,0,blend_radius_m)
  movel([0.292573, -1.406060, -2.547173, -0.759156, 1.570796, 1.863370],accel_mss,speed_ms,0,blend_radius_m)
  movel([0.293532, -1.404124, -2.548612, -0.759653, 1.570796, 1.864328],accel_mss,speed_ms,0,blend_radius_m)
  movel([0.294651, -1.402164, -2.550063, -0.760162, 1.570796, 1.865447],accel_mss,speed_ms,0,blend_radius_m)
  movel([0.295914, -1.400204, -2.551509, -0.760677, 1.570796, 1.866710],accel_mss,speed_ms,0,blend_radius_m)
  movel([0.297300, -1.398268, -2.552930, -0.761191, 1.570796, 1.868097],accel_mss,speed_ms,0,blend_radius_m)
  movel([0.298795, -1.396380, -2.554312, -0.761697, 1.570796, 1.869592],accel_mss,speed_ms,0,blend_radius_m)
  movel([0.300379, -1.394567, -2.555634, -0.762188, 1.570796, 1.871176],accel_mss,speed_ms,0,blend_radius_m)
  movel([0.302032, -1.392854, -2.556878, -0.762657, 1.570796, 1.872828],accel_mss,speed_ms,0,blend_radius_m)
  movel([0.299103, -1.395381, -2.555041, -0.761967, 1.570796, 1.869899],accel_mss,speed_ms,0,blend_radius_m)
  movel([0.296308, -1.398000, -2.553127, -0.761262, 1.570796, 1.867105],accel_mss,speed_ms,0,blend_radius_m)
  movel([0.293641, -1.400694, -2.551147, -0.760547, 1.570796, 1.864437],accel_mss,speed_ms,0,blend_radius_m)
  movel([0.291093, -1.403448, -2.549113, -0.759828, 1.570796, 1.861890],accel_mss,speed_ms,0,blend_radius_m)
  movel([0.288663, -1.406244, -2.547036, -0.759109, 1.570796, 1.859459],accel_mss,speed_ms,0,blend_radius_m)
  movel([0.286339, -1.409068, -2.544927, -0.758394, 1.570796, 1.857136],accel_mss,speed_ms,0,blend_radius_m)
  movel([0.281986, -1.414734, -2.540660, -0.756995, 1.570796, 1.852782],accel_mss,speed_ms,0,blend_radius_m)
  movel([0.283237, -1.412712, -2.542188, -0.757489, 1.570796, 1.854033],accel_mss,speed_ms,0,blend_radius_m)
  movel([0.284296, -1.410491, -2.543860, -0.758038, 1.570796, 1.855093],accel_mss,speed_ms,0,blend_radius_m)
  movel([0.286204, -1.406133, -2.547119, -0.759137, 1.570796, 1.857001],accel_mss,speed_ms,0,blend_radius_m)
  movel([0.287222, -1.404221, -2.548540, -0.759628, 1.570796, 1.858018],accel_mss,speed_ms,0,blend_radius_m)
  movel([0.288274, -1.402524, -2.549797, -0.760068, 1.570796, 1.859070],accel_mss,speed_ms,0,blend_radius_m)
  movel([0.290753, -1.399094, -2.552324, -0.760971, 1.570796, 1.861550],accel_mss,speed_ms,0,blend_radius_m)
  movel([0.290256, -1.399531, -2.552003, -0.760855, 1.570796, 1.861052],accel_mss,speed_ms,0,blend_radius_m)
  movel([0.289438, -1.400025, -2.551640, -0.760724, 1.570796, 1.860235],accel_mss,speed_ms,0,blend_radius_m)
  movel([0.284908, -1.402146, -2.550076, -0.760167, 1.570796, 1.855704],accel_mss,speed_ms,0,blend_radius_m)
  movel([0.283263, -1.402996, -2.549448, -0.759945, 1.570796, 1.854059],accel_mss,speed_ms,0,blend_radius_m)
  movel([0.281380, -1.404403, -2.548405, -0.759581, 1.570796, 1.852176],accel_mss,speed_ms,0,blend_radius_m)
  movel([0.279597, -1.405999, -2.547219, -0.759171, 1.570796, 1.850393],accel_mss,speed_ms,0,blend_radius_m)
  movel([0.276315, -1.409377, -2.544696, -0.758316, 1.570796, 1.847111],accel_mss,speed_ms,0,blend_radius_m)
  movel([0.277669, -1.407465, -2.546126, -0.758798, 1.570796, 1.848465],accel_mss,speed_ms,0,blend_radius_m)
  movel([0.278869, -1.405501, -2.547590, -0.759299, 1.570796, 1.849666],accel_mss,speed_ms,0,blend_radius_m)
  movel([0.281226, -1.401536, -2.550527, -0.760326, 1.570796, 1.852023],accel_mss,speed_ms,0,blend_radius_m)
  movel([0.282639, -1.399519, -2.552012, -0.760858, 1.570796, 1.853435],accel_mss,speed_ms,0,blend_radius_m)
  movel([0.284216, -1.397534, -2.553468, -0.761387, 1.570796, 1.855012],accel_mss,speed_ms,0,blend_radius_m)
  movel([0.287737, -1.393633, -2.556313, -0.762443, 1.570796, 1.858533],accel_mss,speed_ms,0,blend_radius_m)
  movel([0.295224, -1.386069, -2.561766, -0.764554, 1.570796, 1.866020],accel_mss,speed_ms,0,blend_radius_m)
  movel([0.292549, -1.387044, -2.561068, -0.764277, 1.570796, 1.863345],accel_mss,speed_ms,0,blend_radius_m)
  movel([0.289889, -1.388192, -2.560244, -0.763953, 1.570796, 1.860685],accel_mss,speed_ms,0,blend_radius_m)
  movel([0.287257, -1.389501, -2.559302, -0.763586, 1.570796, 1.858053],accel_mss,speed_ms,0,blend_radius_m)
  movel([0.284672, -1.390960, -2.558249, -0.763180, 1.570796, 1.855469],accel_mss,speed_ms,0,blend_radius_m)
  movel([0.282153, -1.392559, -2.557092, -0.762738, 1.570796, 1.852950],accel_mss,speed_ms,0,blend_radius_m)
  movel([0.279712, -1.394290, -2.555835, -0.762264, 1.570796, 1.850509],accel_mss,speed_ms,0,blend_radius_m)
  movel([0.277365, -1.396137, -2.554489, -0.761763, 1.570796, 1.848162],accel_mss,speed_ms,0,blend_radius_m)
  movel([0.275129, -1.398094, -2.553058, -0.761237, 1.570796, 1.845925],accel_mss,speed_ms,0,blend_radius_m)
  movel([0.275734, -1.397461, -2.553522, -0.761407, 1.570796, 1.846531],accel_mss,speed_ms,0,blend_radius_m)
  movel([0.276317, -1.396718, -2.554065, -0.761606, 1.570796, 1.847114],accel_mss,speed_ms,0,blend_radius_m)
  movel([0.277426, -1.395032, -2.555296, -0.762062, 1.570796, 1.848222],accel_mss,speed_ms,0,blend_radius_m)
  movel([0.279464, -1.391765, -2.557668, -0.762957, 1.570796, 1.850260],accel_mss,speed_ms,0,blend_radius_m)
  movel([0.281509, -1.389053, -2.559625, -0.763711, 1.570796, 1.852305],accel_mss,speed_ms,0,blend_radius_m)
  movel([0.283666, -1.386390, -2.561537, -0.764463, 1.570796, 1.854462],accel_mss,speed_ms,0,blend_radius_m)
  movel([0.285930, -1.383774, -2.563404, -0.765211, 1.570796, 1.856726],accel_mss,speed_ms,0,blend_radius_m)
  movel([0.288292, -1.381204, -2.565230, -0.765955, 1.570796, 1.859088],accel_mss,speed_ms,0,blend_radius_m)
  movel([0.290748, -1.378672, -2.567019, -0.766698, 1.570796, 1.861545],accel_mss,speed_ms,0,blend_radius_m)
  movel([0.293295, -1.376180, -2.568772, -0.767438, 1.570796, 1.864091],accel_mss,speed_ms,0,blend_radius_m)
  movel([0.298631, -1.371287, -2.572186, -0.768916, 1.570796, 1.869428],accel_mss,speed_ms,0,blend_radius_m)
  movel([0.296491, -1.372576, -2.571290, -0.768523, 1.570796, 1.867287],accel_mss,speed_ms,0,blend_radius_m)
  movel([0.289931, -1.376010, -2.568891, -0.767488, 1.570796, 1.860727],accel_mss,speed_ms,0,blend_radius_m)
  movel([0.287762, -1.377226, -2.568037, -0.767126, 1.570796, 1.858558],accel_mss,speed_ms,0,blend_radius_m)
  movel([0.285650, -1.378576, -2.567087, -0.766726, 1.570796, 1.856446],accel_mss,speed_ms,0,blend_radius_m)
  movel([0.283665, -1.380083, -2.566023, -0.766283, 1.570796, 1.854461],accel_mss,speed_ms,0,blend_radius_m)
  movel([0.281869, -1.381779, -2.564822, -0.765788, 1.570796, 1.852665],accel_mss,speed_ms,0,blend_radius_m)
  movel([0.284381, -1.378786, -2.566939, -0.766664, 1.570796, 1.855177],accel_mss,speed_ms,0,blend_radius_m)
  movel([0.286891, -1.375635, -2.569153, -0.767600, 1.570796, 1.857687],accel_mss,speed_ms,0,blend_radius_m)
  movel([0.289508, -1.372539, -2.571316, -0.768534, 1.570796, 1.860304],accel_mss,speed_ms,0,blend_radius_m)
  movel([0.290888, -1.371081, -2.572329, -0.768979, 1.570796, 1.861684],accel_mss,speed_ms,0,blend_radius_m)
  movel([0.292335, -1.369721, -2.573272, -0.769396, 1.570796, 1.863131],accel_mss,speed_ms,0,blend_radius_m)
  movel([0.297585, -1.365385, -2.576260, -0.770744, 1.570796, 1.868381],accel_mss,speed_ms,0,blend_radius_m)
  movel([0.302934, -1.361101, -2.579186, -0.772102, 1.570796, 1.873730],accel_mss,speed_ms,0,blend_radius_m)
  movel([0.299202, -1.362838, -2.578003, -0.771548, 1.570796, 1.869998],accel_mss,speed_ms,0,blend_radius_m)
  movel([0.295784, -1.364738, -2.576703, -0.770947, 1.570796, 1.866580],accel_mss,speed_ms,0,blend_radius_m)
  movel([0.292467, -1.366939, -2.575192, -0.770258, 1.570796, 1.863263],accel_mss,speed_ms,0,blend_radius_m)
  movel([0.289040, -1.369569, -2.573377, -0.769443, 1.570796, 1.859836],accel_mss,speed_ms,0,blend_radius_m)
  movel([0.290706, -1.368082, -2.574404, -0.769902, 1.570796, 1.861503],accel_mss,speed_ms,0,blend_radius_m)
  movel([0.292232, -1.366494, -2.575498, -0.770397, 1.570796, 1.863028],accel_mss,speed_ms,0,blend_radius_m)
  movel([0.297867, -1.359716, -2.580127, -0.772546, 1.570796, 1.868664],accel_mss,speed_ms,0,blend_radius_m)
  movel([0.299394, -1.358068, -2.581242, -0.773079, 1.570796, 1.870191],accel_mss,speed_ms,0,blend_radius_m)
  movel([0.301067, -1.356502, -2.582299, -0.773588, 1.570796, 1.871863],accel_mss,speed_ms,0,blend_radius_m)
  movel([0.303440, -1.354630, -2.583557, -0.774201, 1.570796, 1.874236],accel_mss,speed_ms,0,blend_radius_m)
  movel([0.305460, -1.353416, -2.584371, -0.774602, 1.570796, 1.876257],accel_mss,speed_ms,0,blend_radius_m)
  movel([0.305926, -1.353020, -2.584636, -0.774733, 1.570796, 1.876722],accel_mss,speed_ms,0,blend_radius_m)
  movel([0.306116, -1.352575, -2.584934, -0.774880, 1.570796, 1.876912],accel_mss,speed_ms,0,blend_radius_m)
  movel([0.305888, -1.352337, -2.585092, -0.774959, 1.570796, 1.876684],accel_mss,speed_ms,0,blend_radius_m)
  movel([0.305351, -1.352266, -2.585140, -0.774983, 1.570796, 1.876148],accel_mss,speed_ms,0,blend_radius_m)
  movel([0.304613, -1.352325, -2.585101, -0.774963, 1.570796, 1.875409],accel_mss,speed_ms,0,blend_radius_m)
  movel([0.302959, -1.352654, -2.584881, -0.774854, 1.570796, 1.873756],accel_mss,speed_ms,0,blend_radius_m)
  movel([0.301788, -1.353000, -2.584650, -0.774739, 1.570796, 1.872584],accel_mss,speed_ms,0,blend_radius_m)
  movel([0.303760, -1.351220, -2.585838, -0.775331, 1.570796, 1.874556],accel_mss,speed_ms,0,blend_radius_m)
  movel([0.306012, -1.349581, -2.586928, -0.775880, 1.570796, 1.876809],accel_mss,speed_ms,0,blend_radius_m)
  movel([0.310641, -1.346711, -2.588829, -0.776850, 1.570796, 1.881438],accel_mss,speed_ms,0,blend_radius_m)
  speed_ms = 0.005
  movel([0.310641, -1.337928, -2.584667, -0.789794, 1.570796, 1.881438],accel_mss,speed_ms,0,blend_radius_m)
  speed_ms = 0.040
  movel([0.302534, -1.338679, -2.584177, -0.789533, 1.570796, 1.873331],accel_mss,speed_ms,0,blend_radius_m)
  speed_ms = 0.005
  movel([0.302534, -1.347456, -2.588336, -0.776597, 1.570796, 1.873331],accel_mss,speed_ms,0,blend_radius_m)
  speed_ms = 0.025
  movel([0.301969, -1.346437, -2.589009, -0.776943, 1.570796, 1.872765],accel_mss,speed_ms,0,blend_radius_m)
  movel([0.301162, -1.345647, -2.589530, -0.777212, 1.570796, 1.871959],accel_mss,speed_ms,0,blend_radius_m)
  movel([0.300152, -1.345067, -2.589912, -0.777410, 1.570796, 1.870948],accel_mss,speed_ms,0,blend_radius_m)
  movel([0.298976, -1.344675, -2.590170, -0.777545, 1.570796, 1.869773],accel_mss,speed_ms,0,blend_radius_m)
  movel([0.297670, -1.344456, -2.590314, -0.777620, 1.570796, 1.868466],accel_mss,speed_ms,0,blend_radius_m)
  movel([0.296273, -1.344389, -2.590357, -0.777642, 1.570796, 1.867069],accel_mss,speed_ms,0,blend_radius_m)
  movel([0.293350, -1.344628, -2.590200, -0.777560, 1.570796, 1.864146],accel_mss,speed_ms,0,blend_radius_m)
  speed_ms = 0.005
  movel([0.293350, -1.335833, -2.586029, -0.790527, 1.570796, 1.864146],accel_mss,speed_ms,0,blend_radius_m)
  speed_ms = 0.040
  movel([0.305691, -1.331370, -2.588911, -0.792108, 1.570796, 1.876487],accel_mss,speed_ms,0,blend_radius_m)
  speed_ms = 0.005
  movel([0.305691, -1.340193, -2.593102, -0.779094, 1.570796, 1.876487],accel_mss,speed_ms,0,blend_radius_m)
  speed_ms = 0.025
  movel([0.305474, -1.338202, -2.594396, -0.779791, 1.570796, 1.876270],accel_mss,speed_ms,0,blend_radius_m)
  movel([0.305121, -1.336339, -2.595602, -0.780448, 1.570796, 1.875917],accel_mss,speed_ms,0,blend_radius_m)
  movel([0.304577, -1.334650, -2.596691, -0.781048, 1.570796, 1.875373],accel_mss,speed_ms,0,blend_radius_m)
  movel([0.303787, -1.333179, -2.597636, -0.781574, 1.570796, 1.874583],accel_mss,speed_ms,0,blend_radius_m)
  movel([0.302693, -1.331982, -2.598403, -0.782004, 1.570796, 1.873489],accel_mss,speed_ms,0,blend_radius_m)
  movel([0.301247, -1.331099, -2.598968, -0.782322, 1.570796, 1.872043],accel_mss,speed_ms,0,blend_radius_m)
  movel([0.299389, -1.330585, -2.599296, -0.782508, 1.570796, 1.870185],accel_mss,speed_ms,0,blend_radius_m)
  movel([0.298290, -1.330480, -2.599363, -0.782546, 1.570796, 1.869087],accel_mss,speed_ms,0,blend_radius_m)
  movel([0.297068, -1.330485, -2.599360, -0.782544, 1.570796, 1.867865],accel_mss,speed_ms,0,blend_radius_m)
  speed_ms = 0.005
  movel([0.297068, -1.321602, -2.595126, -0.795660, 1.570796, 1.867865],accel_mss,speed_ms,0,blend_radius_m)
  speed_ms = 0.040
  movel([0.307276, -1.318308, -2.597194, -0.796887, 1.570796, 1.878073],accel_mss,speed_ms,0,blend_radius_m)
  speed_ms = 0.005
  movel([0.307276, -1.327210, -2.601442, -0.783736, 1.570796, 1.878073],accel_mss,speed_ms,0,blend_radius_m)
  speed_ms = 0.025
  movel([0.307577, -1.322886, -2.604170, -0.785333, 1.570796, 1.878374],accel_mss,speed_ms,0,blend_radius_m)
  movel([0.307497, -1.320856, -2.605442, -0.786091, 1.570796, 1.878293],accel_mss,speed_ms,0,blend_radius_m)
  movel([0.307183, -1.318969, -2.606619, -0.786801, 1.570796, 1.877979],accel_mss,speed_ms,0,blend_radius_m)
  movel([0.306578, -1.317270, -2.607675, -0.787444, 1.570796, 1.877374],accel_mss,speed_ms,0,blend_radius_m)
  movel([0.305622, -1.315805, -2.608583, -0.788001, 1.570796, 1.876419],accel_mss,speed_ms,0,blend_radius_m)
  movel([0.304256, -1.314613, -2.609319, -0.788457, 1.570796, 1.875052],accel_mss,speed_ms,0,blend_radius_m)
  movel([0.302420, -1.313743, -2.609855, -0.788790, 1.570796, 1.873216],accel_mss,speed_ms,0,blend_radius_m)
  speed_ms = 0.005
  movel([0.302420, -1.304762, -2.605547, -0.802080, 1.570796, 1.873216],accel_mss,speed_ms,0,blend_radius_m)
  speed_ms = 0.040
  movel([0.310889, -1.305667, -2.604996, -0.801726, 1.570796, 1.881685],accel_mss,speed_ms,0,blend_radius_m)
  speed_ms = 0.005
  movel([0.310889, -1.314644, -2.609300, -0.788445, 1.570796, 1.881685],accel_mss,speed_ms,0,blend_radius_m)
  speed_ms = 0.025
  movel([0.311687, -1.311940, -2.610964, -0.789486, 1.570796, 1.882484],accel_mss,speed_ms,0,blend_radius_m)
  movel([0.312325, -1.309202, -2.612638, -0.790549, 1.570796, 1.883121],accel_mss,speed_ms,0,blend_radius_m)
  movel([0.312729, -1.306497, -2.614283, -0.791609, 1.570796, 1.883526],accel_mss,speed_ms,0,blend_radius_m)
  movel([0.312835, -1.303902, -2.615852, -0.792635, 1.570796, 1.883631],accel_mss,speed_ms,0,blend_radius_m)
  movel([0.312571, -1.301486, -2.617305, -0.793598, 1.570796, 1.883367],accel_mss,speed_ms,0,blend_radius_m)
  movel([0.312277, -1.300371, -2.617973, -0.794045, 1.570796, 1.883073],accel_mss,speed_ms,0,blend_radius_m)
  movel([0.311328, -1.298368, -2.619169, -0.794852, 1.570796, 1.882125],accel_mss,speed_ms,0,blend_radius_m)
  movel([0.310655, -1.297501, -2.619685, -0.795203, 1.570796, 1.881451],accel_mss,speed_ms,0,blend_radius_m)
  movel([0.309836, -1.296736, -2.620140, -0.795514, 1.570796, 1.880632],accel_mss,speed_ms,0,blend_radius_m)
  movel([0.308865, -1.296084, -2.620526, -0.795779, 1.570796, 1.879661],accel_mss,speed_ms,0,blend_radius_m)
  speed_ms = 0.005
  movel([0.308865, -1.287004, -2.616138, -0.809246, 1.570796, 1.879661],accel_mss,speed_ms,0,blend_radius_m)
  speed_ms = 0.040
  movel([0.317837, -1.287607, -2.615785, -0.808996, 1.570796, 1.888633],accel_mss,speed_ms,0,blend_radius_m)
  speed_ms = 0.005
  movel([0.317837, -1.296684, -2.620170, -0.795535, 1.570796, 1.888633],accel_mss,speed_ms,0,blend_radius_m)
  speed_ms = 0.025
  movel([0.318956, -1.293496, -2.622056, -0.796836, 1.570796, 1.889753],accel_mss,speed_ms,0,blend_radius_m)
  movel([0.319796, -1.290292, -2.623939, -0.798158, 1.570796, 1.890592],accel_mss,speed_ms,0,blend_radius_m)
  movel([0.320294, -1.287154, -2.625770, -0.799465, 1.570796, 1.891091],accel_mss,speed_ms,0,blend_radius_m)
  movel([0.320374, -1.284175, -2.627497, -0.800718, 1.570796, 1.891171],accel_mss,speed_ms,0,blend_radius_m)
  movel([0.319973, -1.281441, -2.629071, -0.801877, 1.570796, 1.890769],accel_mss,speed_ms,0,blend_radius_m)
  movel([0.319566, -1.280197, -2.629785, -0.802407, 1.570796, 1.890362],accel_mss,speed_ms,0,blend_radius_m)
  movel([0.319015, -1.279047, -2.630442, -0.802900, 1.570796, 1.889812],accel_mss,speed_ms,0,blend_radius_m)
  movel([0.318306, -1.278009, -2.631035, -0.803345, 1.570796, 1.889102],accel_mss,speed_ms,0,blend_radius_m)
  movel([0.317433, -1.277086, -2.631560, -0.803743, 1.570796, 1.888229],accel_mss,speed_ms,0,blend_radius_m)
  movel([0.316387, -1.276300, -2.632007, -0.804082, 1.570796, 1.887183],accel_mss,speed_ms,0,blend_radius_m)
  movel([0.315159, -1.275655, -2.632373, -0.804361, 1.570796, 1.885955],accel_mss,speed_ms,0,blend_radius_m)
  speed_ms = 0.005
  movel([0.315159, -1.266468, -2.627894, -0.818028, 1.570796, 1.885955],accel_mss,speed_ms,0,blend_radius_m)
  speed_ms = 0.040
  movel([0.271584, -1.272863, -2.624289, -0.815237, 1.570796, 1.842380],accel_mss,speed_ms,0,blend_radius_m)
  speed_ms = 0.005
  movel([0.271584, -1.282018, -2.628740, -0.801631, 1.570796, 1.842380],accel_mss,speed_ms,0,blend_radius_m)
  speed_ms = 0.025
  movel([0.273501, -1.283362, -2.627965, -0.801061, 1.570796, 1.844297],accel_mss,speed_ms,0,blend_radius_m)
  movel([0.275155, -1.284971, -2.627036, -0.800382, 1.570796, 1.845952],accel_mss,speed_ms,0,blend_radius_m)
  movel([0.276562, -1.286817, -2.625966, -0.799606, 1.570796, 1.847358],accel_mss,speed_ms,0,blend_radius_m)
  movel([0.277730, -1.288874, -2.624768, -0.798747, 1.570796, 1.848527],accel_mss,speed_ms,0,blend_radius_m)
  movel([0.278667, -1.291117, -2.623455, -0.797817, 1.570796, 1.849463],accel_mss,speed_ms,0,blend_radius_m)
  movel([0.279390, -1.293520, -2.622042, -0.796827, 1.570796, 1.850186],accel_mss,speed_ms,0,blend_radius_m)
  movel([0.279902, -1.296060, -2.620540, -0.795788, 1.570796, 1.850698],accel_mss,speed_ms,0,blend_radius_m)
  movel([0.280222, -1.298709, -2.618966, -0.794714, 1.570796, 1.851018],accel_mss,speed_ms,0,blend_radius_m)
  movel([0.280353, -1.301443, -2.617331, -0.793615, 1.570796, 1.851149],accel_mss,speed_ms,0,blend_radius_m)
  movel([0.280314, -1.304241, -2.615648, -0.792501, 1.570796, 1.851110],accel_mss,speed_ms,0,blend_radius_m)
  movel([0.280111, -1.307074, -2.613933, -0.791382, 1.570796, 1.850907],accel_mss,speed_ms,0,blend_radius_m)
  movel([0.279756, -1.309927, -2.612196, -0.790266, 1.570796, 1.850552],accel_mss,speed_ms,0,blend_radius_m)
  movel([0.279261, -1.312769, -2.610455, -0.789166, 1.570796, 1.850057],accel_mss,speed_ms,0,blend_radius_m)
  movel([0.278632, -1.315586, -2.608718, -0.788085, 1.570796, 1.849428],accel_mss,speed_ms,0,blend_radius_m)
  movel([0.277883, -1.318348, -2.607006, -0.787035, 1.570796, 1.848680],accel_mss,speed_ms,0,blend_radius_m)
  movel([0.277026, -1.321040, -2.605327, -0.786022, 1.570796, 1.847823],accel_mss,speed_ms,0,blend_radius_m)
  movel([0.275722, -1.324606, -2.603088, -0.784695, 1.570796, 1.846518],accel_mss,speed_ms,0,blend_radius_m)
  movel([0.274014, -1.328675, -2.600512, -0.783201, 1.570796, 1.844810],accel_mss,speed_ms,0,blend_radius_m)
  movel([0.271907, -1.332885, -2.597825, -0.781679, 1.570796, 1.842703],accel_mss,speed_ms,0,blend_radius_m)
  movel([0.270705, -1.334932, -2.596509, -0.780948, 1.570796, 1.841501],accel_mss,speed_ms,0,blend_radius_m)
  movel([0.269409, -1.336880, -2.595252, -0.780257, 1.570796, 1.840206],accel_mss,speed_ms,0,blend_radius_m)
  movel([0.268012, -1.338693, -2.594077, -0.779619, 1.570796, 1.838808],accel_mss,speed_ms,0,blend_radius_m)
  movel([0.266519, -1.340319, -2.593020, -0.779050, 1.570796, 1.837315],accel_mss,speed_ms,0,blend_radius_m)
  movel([0.264925, -1.341725, -2.592103, -0.778561, 1.570796, 1.835721],accel_mss,speed_ms,0,blend_radius_m)
  movel([0.263229, -1.342867, -2.591356, -0.778166, 1.570796, 1.834025],accel_mss,speed_ms,0,blend_radius_m)
  movel([0.261433, -1.343701, -2.590809, -0.777879, 1.570796, 1.832229],accel_mss,speed_ms,0,blend_radius_m)
  movel([0.259532, -1.344191, -2.590487, -0.777710, 1.570796, 1.830328],accel_mss,speed_ms,0,blend_radius_m)
  movel([0.258540, -1.344293, -2.590421, -0.777676, 1.570796, 1.829336],accel_mss,speed_ms,0,blend_radius_m)
  movel([0.257520, -1.344293, -2.590421, -0.777676, 1.570796, 1.828316],accel_mss,speed_ms,0,blend_radius_m)
  movel([0.255398, -1.343965, -2.590636, -0.777788, 1.570796, 1.826194],accel_mss,speed_ms,0,blend_radius_m)
  movel([0.253024, -1.343213, -2.591129, -0.778047, 1.570796, 1.823820],accel_mss,speed_ms,0,blend_radius_m)
  movel([0.250895, -1.342245, -2.591763, -0.778381, 1.570796, 1.821691],accel_mss,speed_ms,0,blend_radius_m)
  movel([0.248983, -1.341083, -2.592522, -0.778784, 1.570796, 1.819779],accel_mss,speed_ms,0,blend_radius_m)
  movel([0.247251, -1.339740, -2.593397, -0.779252, 1.570796, 1.818048],accel_mss,speed_ms,0,blend_radius_m)
  movel([0.245674, -1.338235, -2.594374, -0.779779, 1.570796, 1.816470],accel_mss,speed_ms,0,blend_radius_m)
  movel([0.244216, -1.336590, -2.595440, -0.780360, 1.570796, 1.815012],accel_mss,speed_ms,0,blend_radius_m)
  movel([0.241528, -1.332939, -2.597790, -0.781660, 1.570796, 1.812324],accel_mss,speed_ms,0,blend_radius_m)
  movel([0.238720, -1.328765, -2.600456, -0.783169, 1.570796, 1.809516],accel_mss,speed_ms,0,blend_radius_m)
  movel([0.236045, -1.324512, -2.603147, -0.784730, 1.570796, 1.806841],accel_mss,speed_ms,0,blend_radius_m)
  movel([0.233638, -1.320040, -2.605952, -0.786398, 1.570796, 1.804435],accel_mss,speed_ms,0,blend_radius_m)
  movel([0.232584, -1.317672, -2.607426, -0.787291, 1.570796, 1.803380],accel_mss,speed_ms,0,blend_radius_m)
  movel([0.231653, -1.315190, -2.608963, -0.788236, 1.570796, 1.802449],accel_mss,speed_ms,0,blend_radius_m)
  movel([0.230440, -1.312125, -2.610850, -0.789414, 1.570796, 1.801236],accel_mss,speed_ms,0,blend_radius_m)
  movel([0.228947, -1.309165, -2.612660, -0.790563, 1.570796, 1.799743],accel_mss,speed_ms,0,blend_radius_m)
  movel([0.227212, -1.306316, -2.614393, -0.791680, 1.570796, 1.798008],accel_mss,speed_ms,0,blend_radius_m)
  movel([0.225283, -1.303570, -2.616052, -0.792767, 1.570796, 1.796079],accel_mss,speed_ms,0,blend_radius_m)
  movel([0.221008, -1.298396, -2.619152, -0.794841, 1.570796, 1.791805],accel_mss,speed_ms,0,blend_radius_m)
  movel([0.216480, -1.293618, -2.621985, -0.796787, 1.570796, 1.787276],accel_mss,speed_ms,0,blend_radius_m)
  movel([0.212807, -1.290271, -2.623951, -0.798167, 1.570796, 1.783603],accel_mss,speed_ms,0,blend_radius_m)
  movel([0.208744, -1.287288, -2.625692, -0.799409, 1.570796, 1.779540],accel_mss,speed_ms,0,blend_radius_m)
  movel([0.204297, -1.284701, -2.627192, -0.800496, 1.570796, 1.775094],accel_mss,speed_ms,0,blend_radius_m)
  movel([0.199477, -1.282551, -2.628433, -0.801405, 1.570796, 1.770273],accel_mss,speed_ms,0,blend_radius_m)
  movel([0.194294, -1.280863, -2.629403, -0.802123, 1.570796, 1.765090],accel_mss,speed_ms,0,blend_radius_m)
  movel([0.191571, -1.280203, -2.629781, -0.802405, 1.570796, 1.762368],accel_mss,speed_ms,0,blend_radius_m)
  movel([0.185870, -1.279270, -2.630315, -0.802804, 1.570796, 1.756666],accel_mss,speed_ms,0,blend_radius_m)
  movel([0.182894, -1.279004, -2.630467, -0.802918, 1.570796, 1.753690],accel_mss,speed_ms,0,blend_radius_m)
  movel([0.176709, -1.278890, -2.630532, -0.802967, 1.570796, 1.747505],accel_mss,speed_ms,0,blend_radius_m)
  movel([0.172314, -1.279205, -2.630352, -0.802832, 1.570796, 1.743111],accel_mss,speed_ms,0,blend_radius_m)
  movel([0.167777, -1.279921, -2.629943, -0.802525, 1.570796, 1.738574],accel_mss,speed_ms,0,blend_radius_m)
  movel([0.163141, -1.281034, -2.629305, -0.802050, 1.570796, 1.733937],accel_mss,speed_ms,0,blend_radius_m)
  movel([0.158445, -1.282545, -2.628437, -0.801408, 1.570796, 1.729241],accel_mss,speed_ms,0,blend_radius_m)
  movel([0.153727, -1.284450, -2.627337, -0.800602, 1.570796, 1.724524],accel_mss,speed_ms,0,blend_radius_m)
  movel([0.149032, -1.286744, -2.626008, -0.799637, 1.570796, 1.719828],accel_mss,speed_ms,0,blend_radius_m)
  movel([0.144398, -1.289420, -2.624449, -0.798520, 1.570796, 1.715194],accel_mss,speed_ms,0,blend_radius_m)
  movel([0.139866, -1.292470, -2.622660, -0.797258, 1.570796, 1.710662],accel_mss,speed_ms,0,blend_radius_m)
  movel([0.135776, -1.295589, -2.620820, -0.795980, 1.570796, 1.706572],accel_mss,speed_ms,0,blend_radius_m)
  movel([0.131973, -1.298825, -2.618896, -0.794667, 1.570796, 1.702770],accel_mss,speed_ms,0,blend_radius_m)
  movel([0.128482, -1.302183, -2.616887, -0.793319, 1.570796, 1.699278],accel_mss,speed_ms,0,blend_radius_m)
